// Core 3.10.2: deterministic typed walk, one bounded response window.
// Static facets carry no write capability. Every reused slot is cleared.
FUNCTION "FRK_ConfigRevision" : UDInt
{ S7_Optimized_Access := 'TRUE' }
VERSION : 0.1
VAR_INPUT
    Previous : UDInt;
END_VAR
VAR_TEMP
    Stamp : DTL;
    ResultCode : Int;
    Generation : ULInt;
END_VAR
BEGIN
    #FRK_ConfigRevision := #Previous + 1;
    #ResultCode := RD_SYS_T(OUT => #Stamp);
    IF #ResultCode = 0 THEN
        #Generation := LDT_TO_ULINT(DTL_TO_LDT(#Stamp)) / ULINT#1000000;
        #FRK_ConfigRevision := ULINT_TO_UDINT(#Generation MOD ULINT#4294967296);
    END_IF;
    IF #FRK_ConfigRevision = #Previous THEN #FRK_ConfigRevision := #Previous + 1; END_IF;
    IF #FRK_ConfigRevision = 0 THEN #FRK_ConfigRevision := 1; END_IF;
END_FUNCTION

FUNCTION "FRK_ConfigBegin" : Void
{ S7_Optimized_Access := 'TRUE' }
VERSION : 0.1
VAR_INPUT
    PageIndex : DInt;
    Revision : UDInt;
END_VAR
VAR_IN_OUT
    Cursor : "FRK_ConfigCursor";
    Page : "ST_ConfigPage";
END_VAR
VAR_TEMP
    Index : Int;
END_VAR
BEGIN
    #Cursor.Position := 0;
    #Cursor.First := 0;
    #Page.Revision := #Revision;
    #Page.PageIndex := 0;
    IF #PageIndex >= 0 AND #PageIndex <= 32767 THEN
        #Cursor.First := #PageIndex * 16;
        #Page.PageIndex := DINT_TO_INT(#PageIndex);
    END_IF;
    #Page.PageCount := 1;
    #Page.EntryCount := 0;
    "FRK_UnitScratch".EmptyConfigEntry.ValueType := 1;
    "FRK_UnitScratch".EmptyConfigEntry.Readable := TRUE;
    FOR #Index := 1 TO 16 DO
        #Page.Entries[#Index] := "FRK_UnitScratch".EmptyConfigEntry;
    END_FOR;
END_FUNCTION

FUNCTION "FRK_ConfigAppend" : Void
{ S7_Optimized_Access := 'TRUE' }
VERSION : 0.1
VAR_INPUT
    Scope : String;
    Item : String;
    ValueText : WString;
    ValueType : DInt;
    ReadLevel : DInt;
    Readable : Bool;
END_VAR
VAR_IN_OUT
    Cursor : "FRK_ConfigCursor";
    Page : "ST_ConfigPage";
END_VAR
VAR_TEMP
    Slot : DInt;
END_VAR
BEGIN
    #Slot := #Cursor.Position - #Cursor.First;
    #Cursor.Position := #Cursor.Position + 1;
    IF #Slot < 0 OR #Slot >= 16 THEN RETURN; END_IF;
    #Slot := #Slot + 1;
    #Page.Entries[#Slot].Scope := STRING_TO_WSTRING(#Scope);
    #Page.Entries[#Slot].Item := STRING_TO_WSTRING(#Item);
    #Page.Entries[#Slot].ValueType := #ValueType;
    #Page.Entries[#Slot].ReadLevel := #ReadLevel;
    #Page.Entries[#Slot].Readable := #Readable;
    IF #Readable THEN #Page.Entries[#Slot].ValueText := #ValueText; END_IF;
    #Page.EntryCount := DINT_TO_INT(#Slot);
END_FUNCTION

FUNCTION "FRK_ConfigFinish" : Void
{ S7_Optimized_Access := 'TRUE' }
VERSION : 0.1
VAR_IN_OUT
    Cursor : "FRK_ConfigCursor";
    Page : "ST_ConfigPage";
END_VAR
BEGIN
    #Page.PageCount := DINT_TO_INT((#Cursor.Position + 16 - 1) / 16);
    IF #Page.PageCount < 1 THEN #Page.PageCount := 1; END_IF;
END_FUNCTION

FUNCTION "FRK_ConfigCatalog" : Void
{ S7_Optimized_Access := 'TRUE' }
VERSION : 0.1
VAR_INPUT
    Scope : String;
    Count : Int;
    Catalog : Array[1..12] of "ST_CommandInfo";
    ReadLevel : DInt;
    Readable : Bool;
END_VAR
VAR_IN_OUT
    Cursor : "FRK_ConfigCursor";
    Page : "ST_ConfigPage";
END_VAR
VAR_TEMP
    Index : Int;
    IndexText : String[8];
    Prefix : String[254];
    Item : String[254];
END_VAR
BEGIN
    "FRK_ConfigAppend"(Scope := #Scope, Item := 'CatalogCount', ValueText := STRING_TO_WSTRING(INT_TO_STRING(#Count)), ValueType := 0, ReadLevel := #ReadLevel, Readable := #Readable, Cursor := #Cursor, Page := #Page);
    FOR #Index := 1 TO #Count DO
        IF #Index > 12 THEN EXIT; END_IF;
        #IndexText := INT_TO_STRING(#Index);
        IF #IndexText[1] = '+' THEN #IndexText := DELETE(IN := #IndexText, L := 1, P := 1); END_IF;
        #Prefix := CONCAT(IN1 := 'Catalog/Catalog[', IN2 := #IndexText);
        #Prefix := CONCAT(IN1 := #Prefix, IN2 := ']/');
        #Item := CONCAT(IN1 := #Prefix, IN2 := 'Value');
        "FRK_ConfigAppend"(Scope := #Scope, Item := #Item, ValueText := STRING_TO_WSTRING(DINT_TO_STRING(#Catalog[#Index].Value)), ValueType := 0, ReadLevel := #ReadLevel, Readable := #Readable, Cursor := #Cursor, Page := #Page);
        #Item := CONCAT(IN1 := #Prefix, IN2 := 'Label');
        "FRK_ConfigAppend"(Scope := #Scope, Item := #Item, ValueText := STRING_TO_WSTRING(#Catalog[#Index].Label), ValueType := 1, ReadLevel := #ReadLevel, Readable := #Readable, Cursor := #Cursor, Page := #Page);
        #Item := CONCAT(IN1 := #Prefix, IN2 := 'Style');
        "FRK_ConfigAppend"(Scope := #Scope, Item := #Item, ValueText := STRING_TO_WSTRING(DINT_TO_STRING(#Catalog[#Index].Style)), ValueType := 0, ReadLevel := #ReadLevel, Readable := #Readable, Cursor := #Cursor, Page := #Page);
    END_FOR;
END_FUNCTION

FUNCTION "FRK_ConfigUnit" : Void
{ S7_Optimized_Access := 'TRUE' }
VERSION : 0.1
VAR_INPUT
    Scope : String;
    Policy : Array[0..6] of "ST_ModePolicy";
    ModelCount : Int;
    ReadLevel : DInt;
    Readable : Bool;
END_VAR
VAR_IN_OUT
    Cursor : "FRK_ConfigCursor";
    Page : "ST_ConfigPage";
END_VAR
VAR_TEMP
    Index : Int;
    IndexText : String[8];
    Prefix : String[254];
    Item : String[254];
END_VAR
BEGIN
    "FRK_ConfigAppend"(Scope := #Scope, Item := 'CatalogCount', ValueText := WSTRING#'0', ValueType := 0, ReadLevel := #ReadLevel, Readable := #Readable, Cursor := #Cursor, Page := #Page);
    "FRK_ConfigAppend"(Scope := #Scope, Item := 'AvailableModelCount', ValueText := INT_TO_WSTRING(#ModelCount), ValueType := 0, ReadLevel := #ReadLevel, Readable := #Readable, Cursor := #Cursor, Page := #Page);
    FOR #Index := 0 TO 6 DO
        #IndexText := INT_TO_STRING(#Index);
        IF #IndexText[1] = '+' THEN #IndexText := DELETE(IN := #IndexText, L := 1, P := 1); END_IF;
        #Prefix := CONCAT(IN1 := 'ModePolicy/ModePolicy[', IN2 := #IndexText);
        #Prefix := CONCAT(IN1 := #Prefix, IN2 := ']/');
        #Item := CONCAT(IN1 := #Prefix, IN2 := 'Shield');
        "FRK_ConfigAppend"(Scope := #Scope, Item := #Item, ValueText := STRING_TO_WSTRING(DINT_TO_STRING(#Policy[#Index].Shield)), ValueType := 0, ReadLevel := #ReadLevel, Readable := #Readable, Cursor := #Cursor, Page := #Page);
        #Item := CONCAT(IN1 := #Prefix, IN2 := 'Style');
        "FRK_ConfigAppend"(Scope := #Scope, Item := #Item, ValueText := STRING_TO_WSTRING(DINT_TO_STRING(#Policy[#Index].Style)), ValueType := 0, ReadLevel := #ReadLevel, Readable := #Readable, Cursor := #Cursor, Page := #Page);
    END_FOR;
END_FUNCTION

// Core 8.3: one owning active list / closed ring, with optional event callback.
FUNCTION "FRK_AlarmNotify" : Void
{ S7_Optimized_Access := 'TRUE' }
VERSION : 0.1
VAR_INPUT
    Ev : "ST_AlarmEvent";
END_VAR
VAR_IN_OUT
    AlarmLog : "FRK_AlarmLog";
END_VAR
BEGIN
    RETURN; // No event sink supplied by the composition declaration.
END_FUNCTION

FUNCTION "FRK_AlarmRefresh" : Void
{ S7_Optimized_Access := 'TRUE' }
VERSION : 0.1
VAR_IN_OUT
    AlarmLog : "FRK_AlarmLog";
END_VAR
VAR_TEMP
    Index : Int;
END_VAR
BEGIN
    #AlarmLog.NActive := 0;
    #AlarmLog.Blocking := FALSE;
    FOR #Index := 1 TO 16 DO
        IF #AlarmLog.Active[#Index].State <> 0 THEN
            #AlarmLog.NActive := #AlarmLog.NActive + 1;
            IF #AlarmLog.Active[#Index].ResetClass = 1 THEN #AlarmLog.Blocking := TRUE; END_IF;
        END_IF;
    END_FOR;
    "FRK_AlarmRecoveryRefresh"(AlarmLog := #AlarmLog);
END_FUNCTION

FUNCTION "FRK_AlarmBegin" : Void
{ S7_Optimized_Access := 'TRUE' }
VERSION : 0.1
VAR_INPUT
    Startup : Bool;
END_VAR
VAR_IN_OUT
    AlarmLog : "FRK_AlarmLog";
END_VAR
VAR_TEMP
    Index : Int;
END_VAR
BEGIN
    FOR #Index := 1 TO 16 DO
        #AlarmLog.Touched[#Index] := FALSE;
        IF #Startup THEN
            #AlarmLog.Active[#Index] := "FRK_UnitScratch".EmptyEvent;
            #AlarmLog.Automatic[#Index] := FALSE;
            #AlarmLog.ComeMs[#Index] := 0;
        END_IF;
    END_FOR;
    IF #Startup THEN
        FOR #Index := 1 TO 64 DO #AlarmLog.Ring[#Index] := "FRK_UnitScratch".EmptyEvent; END_FOR;
        #AlarmLog.RingHead := 0;
        #AlarmLog.RingUsed := 0;
        #AlarmLog.Truncated := FALSE;
    END_IF;
    IF #Startup AND #AlarmLog.HistorySlot > 0 THEN "FRK_AlarmHistoryClear"(AlarmLog := #AlarmLog); END_IF;
    IF #Startup THEN "FRK_AlarmRecoveryClear"(AlarmLog := #AlarmLog); END_IF;
    "FRK_AlarmRefresh"(AlarmLog := #AlarmLog);
END_FUNCTION

FUNCTION "FRK_AlarmRaise" : Int
{ S7_Optimized_Access := 'TRUE' }
VERSION : 0.1
VAR_INPUT
    Diag : "ST_Diagnostic";
    ResetClass : DInt;
END_VAR
VAR_IN_OUT
    AlarmLog : "FRK_AlarmLog";
END_VAR
VAR_TEMP
    Slot : Int;
    Stamp : DTL;
    ResultCode : Int;
    Rational : "ST_Diagnostic";
END_VAR
BEGIN
    #FRK_AlarmRaise := 0;
    IF #ResetClass < 0 OR #ResetClass > 1
        OR #Diag.Severity < 0 OR #Diag.Severity > 2
        OR #Diag.Category < 0 OR #Diag.Category > 2
        OR #Diag.SourcePath = WSTRING#'' OR #Diag.Description = WSTRING#'' THEN RETURN; END_IF;
    #Slot := "FRK_AlarmRecoveryClaim"(AlarmLog := #AlarmLog, Diag := #Diag, ResetClass := #ResetClass); IF #Slot > 0 THEN #FRK_AlarmRaise := #Slot; RETURN; END_IF;
    FOR #Slot := 1 TO 16 DO
        IF #AlarmLog.Active[#Slot].State = 0 THEN
            #Rational := #Diag;
            "FRK_Rationalize"(Diag := #Rational);
            #AlarmLog.Active[#Slot] := "FRK_UnitScratch".EmptyEvent;
            #AlarmLog.Active[#Slot].ReasonCode := #Rational.ReasonCode;
            #AlarmLog.Active[#Slot].Description := #Rational.Description;
            #AlarmLog.Active[#Slot].SourcePath := #Rational.SourcePath;
            #AlarmLog.Active[#Slot].IoTag := #Rational.IoTag;
            #AlarmLog.Active[#Slot].IoAddress := #Rational.IoAddress;
            #AlarmLog.Active[#Slot].Severity := #Rational.Severity;
            #AlarmLog.Active[#Slot].Category := #Rational.Category;
            #AlarmLog.Active[#Slot].ResetClass := #ResetClass;
            #AlarmLog.Active[#Slot].State := 1;
            #AlarmLog.ComeMs[#Slot] := "FRK_Clock".NowMs;
            #AlarmLog.ElapsedBefore[#Slot] := 0; #AlarmLog.Recovering[#Slot] := FALSE;
            #AlarmLog.Automatic[#Slot] := FALSE;
            #AlarmLog.Touched[#Slot] := FALSE;
            #ResultCode := RD_SYS_T(OUT => #Stamp);
            IF #ResultCode = 0 THEN #AlarmLog.Active[#Slot].ComeAt := DTL_TO_LDT(#Stamp); END_IF;
            // The UTC source has no proven synchronization witness yet.
            #AlarmLog.Active[#Slot].ComeTimeSynchronized := FALSE;
            "FRK_AlarmRefresh"(AlarmLog := #AlarmLog);
            "FRK_AlarmRecoveryStore"(AlarmLog := #AlarmLog, EventSlot := #Slot);
            "FRK_DeliveryCapture"(AlarmLog := #AlarmLog, Ev := #AlarmLog.Active[#Slot]);
            "FRK_AlarmNotify"(AlarmLog := #AlarmLog, Ev := #AlarmLog.Active[#Slot]);
            #FRK_AlarmRaise := #Slot;
            RETURN;
        END_IF;
    END_FOR;
    IF NOT #AlarmLog.Truncated THEN
        #AlarmLog.Truncated := TRUE;
        "FRK_AlarmHistoryHeaderSave"(AlarmLog := #AlarmLog);
    END_IF;
END_FUNCTION

FUNCTION "FRK_AlarmClose" : Void
{ S7_Optimized_Access := 'TRUE' }
VERSION : 0.1
VAR_INPUT
    Slot : Int;
END_VAR
VAR_IN_OUT
    AlarmLog : "FRK_AlarmLog";
END_VAR
BEGIN
    IF #Slot < 1 OR #Slot > 16 THEN RETURN; END_IF;
    IF #AlarmLog.Active[#Slot].State = 0 THEN RETURN; END_IF;
    #AlarmLog.Active[#Slot].State := 0;
    "FRK_DeliveryCapture"(AlarmLog := #AlarmLog, Ev := #AlarmLog.Active[#Slot]);
    "FRK_AlarmRecoveryClosePrepare"(AlarmLog := #AlarmLog, EventSlot := #Slot);
    IF #AlarmLog.RingHead < 0 OR #AlarmLog.RingHead > 64 THEN #AlarmLog.RingHead := 0; END_IF;
    #AlarmLog.RingHead := (#AlarmLog.RingHead MOD 64) + 1;
    IF #AlarmLog.RingUsed >= 64 THEN #AlarmLog.Truncated := TRUE;
    ELSE #AlarmLog.RingUsed := #AlarmLog.RingUsed + 1; END_IF;
    #AlarmLog.Ring[#AlarmLog.RingHead] := #AlarmLog.Active[#Slot];
    "FRK_AlarmHistoryAppend"(AlarmLog := #AlarmLog);
    "FRK_AlarmRecoveryStore"(AlarmLog := #AlarmLog, EventSlot := #Slot);
    #AlarmLog.Automatic[#Slot] := FALSE;
    "FRK_AlarmRefresh"(AlarmLog := #AlarmLog);
    "FRK_AlarmNotify"(AlarmLog := #AlarmLog, Ev := #AlarmLog.Ring[#AlarmLog.RingHead]);
END_FUNCTION

FUNCTION "FRK_AlarmGone" : Bool
{ S7_Optimized_Access := 'TRUE' }
VERSION : 0.1
VAR_INPUT
    Slot : Int;
END_VAR
VAR_IN_OUT
    AlarmLog : "FRK_AlarmLog";
END_VAR
VAR_TEMP
    Span : UDInt;
    Stamp : DTL;
    ResultCode : Int;
END_VAR
BEGIN
    #FRK_AlarmGone := FALSE;
    IF #Slot < 1 OR #Slot > 16 THEN RETURN; END_IF;
    IF #AlarmLog.Active[#Slot].State <> 1 THEN RETURN; END_IF;
    #ResultCode := RD_SYS_T(OUT => #Stamp);
    IF #ResultCode = 0 THEN #AlarmLog.Active[#Slot].GoneAt := DTL_TO_LDT(#Stamp); END_IF;
    #AlarmLog.Active[#Slot].GoneTimeSynchronized := FALSE;
    #Span := "FRK_AlarmRecoveryElapsed"(AlarmLog := #AlarmLog, EventSlot := #Slot);
    #AlarmLog.Active[#Slot].Duration := DINT_TO_TIME(UDINT_TO_DINT(#Span));
    IF #AlarmLog.Active[#Slot].ResetClass = 0 THEN
        "FRK_AlarmClose"(AlarmLog := #AlarmLog, Slot := #Slot);
    ELSE
        #AlarmLog.Active[#Slot].State := 2;
        #AlarmLog.Automatic[#Slot] := FALSE;
        "FRK_AlarmRecoveryStore"(AlarmLog := #AlarmLog, EventSlot := #Slot);
    END_IF;
    #FRK_AlarmGone := TRUE;
END_FUNCTION

FUNCTION "FRK_AlarmOperatorReset" : Void
{ S7_Optimized_Access := 'TRUE' }
VERSION : 0.1
VAR_IN_OUT
    AlarmLog : "FRK_AlarmLog";
END_VAR
VAR_TEMP
    Slot : Int;
    Gone : Bool;
    Stamp : DTL;
    ResultCode : Int;
END_VAR
BEGIN
    FOR #Slot := 1 TO 16 DO
        IF #AlarmLog.Active[#Slot].State <> 0 AND #AlarmLog.Active[#Slot].ResetClass = 1 THEN
            IF #AlarmLog.Active[#Slot].State = 1 THEN #Gone := "FRK_AlarmGone"(AlarmLog := #AlarmLog, Slot := #Slot); END_IF;
            #ResultCode := RD_SYS_T(OUT => #Stamp);
            IF #ResultCode = 0 THEN #AlarmLog.Active[#Slot].ResetAt := DTL_TO_LDT(#Stamp); END_IF;
            #AlarmLog.Active[#Slot].ResetTimeSynchronized := FALSE;
            "FRK_AlarmClose"(AlarmLog := #AlarmLog, Slot := #Slot);
        END_IF;
    END_FOR;
END_FUNCTION

FUNCTION "FRK_AlarmMessage" : Void
{ S7_Optimized_Access := 'TRUE' }
VERSION : 0.1
VAR_INPUT
    Reason : DInt;
    Description : WString;
    SourcePath : WString;
END_VAR
VAR_IN_OUT
    AlarmLog : "FRK_AlarmLog";
END_VAR
VAR_TEMP
    Diag : "ST_Diagnostic";
    Slot : Int;
    Gone : Bool;
END_VAR
BEGIN
    #Diag := "FRK_UnitScratch".EmptyDiagnostic;
    #Diag.ReasonCode := #Reason;
    #Diag.Description := #Description;
    #Diag.SourcePath := #SourcePath;
    #Diag.Severity := 0;
    #Diag.Category := 2;
    #Slot := "FRK_AlarmRaise"(AlarmLog := #AlarmLog, Diag := #Diag, ResetClass := 0);
    IF #Slot > 0 THEN #Gone := "FRK_AlarmGone"(AlarmLog := #AlarmLog, Slot := #Slot); END_IF;
END_FUNCTION

FUNCTION "FRK_AlarmCapture" : Void
{ S7_Optimized_Access := 'TRUE' }
VERSION : 0.1
VAR_IN_OUT
    AlarmLog : "FRK_AlarmLog";
    Core : "FRK_Core";
    Status : "ST_ModuleStatus";
END_VAR
VAR_TEMP
    Slot : Int;
END_VAR
BEGIN
    #Slot := #Core.FaultSlot;
    IF #Slot < 1 OR #Slot > 16 THEN #Slot := 0;
    ELSIF NOT #AlarmLog.Automatic[#Slot] OR #AlarmLog.Active[#Slot].State <> 1
        OR #AlarmLog.Active[#Slot].SourcePath <> #Status.Diagnostic.SourcePath
        OR #AlarmLog.Active[#Slot].ReasonCode <> #Status.Diagnostic.ReasonCode
        OR #AlarmLog.Active[#Slot].Description <> #Status.Diagnostic.Description THEN #Slot := 0; END_IF;
    IF #Core.Exec = 3 AND NOT #Core.FaultHandled THEN
        IF #Slot = 0 THEN
            // Adopted first-outs share one active occurrence within this log.
            FOR #Slot := 1 TO 16 DO
                IF #AlarmLog.Automatic[#Slot] AND #AlarmLog.Active[#Slot].State = 1
                    AND #AlarmLog.Active[#Slot].SourcePath = #Status.Diagnostic.SourcePath
                    AND #AlarmLog.Active[#Slot].ReasonCode = #Status.Diagnostic.ReasonCode
                    AND #AlarmLog.Active[#Slot].Description = #Status.Diagnostic.Description THEN EXIT; END_IF;
            END_FOR;
            IF #Slot > 16 THEN #Slot := "FRK_AlarmRaise"(AlarmLog := #AlarmLog, Diag := #Status.Diagnostic, ResetClass := 1); END_IF;
        END_IF;
        IF #Slot > 0 THEN IF NOT #AlarmLog.Automatic[#Slot] THEN #AlarmLog.Automatic[#Slot] := TRUE; "FRK_AlarmRecoveryStore"(AlarmLog := #AlarmLog, EventSlot := #Slot); END_IF; #AlarmLog.Recovering[#Slot] := FALSE; #AlarmLog.Automatic[#Slot] := TRUE; #AlarmLog.Touched[#Slot] := TRUE; END_IF;
        #Core.FaultSlot := #Slot;
    ELSE
        #Core.FaultSlot := 0;
    END_IF;
END_FUNCTION

FUNCTION "FRK_AlarmEnd" : Void
{ S7_Optimized_Access := 'TRUE' }
VERSION : 0.1
VAR_IN_OUT
    AlarmLog : "FRK_AlarmLog";
END_VAR
VAR_TEMP
    Slot : Int;
    Gone : Bool;
END_VAR
BEGIN
    FOR #Slot := 1 TO 16 DO
        IF #AlarmLog.Automatic[#Slot] AND NOT #AlarmLog.Touched[#Slot] THEN #Gone := "FRK_AlarmGone"(AlarmLog := #AlarmLog, Slot := #Slot); END_IF;
    END_FOR;
END_FUNCTION

FUNCTION "FRK_AlarmTreeBlocking" : Bool
{ S7_Optimized_Access := 'TRUE' }
VERSION : 0.1
VAR_INPUT
    Owner : DInt;
END_VAR
VAR_TEMP
    Index : DInt;
    Ancestor : DInt;
    Depth : DInt;
END_VAR
BEGIN
    #FRK_AlarmTreeBlocking := TRUE;
    IF "FRK_Registry".Fault OR #Owner < 1 OR #Owner > "FRK_Registry".Count OR "FRK_Registry".Count > 4 THEN RETURN; END_IF;
    FOR #Index := 1 TO "FRK_Registry".Count DO
        IF "FRK_Registry".Rows[#Index].AlarmBlocking THEN
            #Ancestor := #Index;
            FOR #Depth := 1 TO 4 DO
                IF #Ancestor = #Owner THEN RETURN; END_IF;
                IF #Ancestor = 0 THEN EXIT; END_IF;
                IF #Ancestor < 1 OR #Ancestor > "FRK_Registry".Count THEN RETURN; END_IF;
                #Ancestor := "FRK_Registry".Rows[#Ancestor].Parent;
            END_FOR;
            IF #Depth > 4 AND #Ancestor <> 0 THEN RETURN; END_IF;
        END_IF;
    END_FOR;
    #FRK_AlarmTreeBlocking := FALSE;
END_FUNCTION

// Reference-1500 LOCAL_RETAIN: closed history only, keyed by actual Unit scope.
// No active alarms, commands, sessions or monotonic clocks are restored.
FUNCTION "FRK_AlarmHistoryIndex" : Int
{ S7_Optimized_Access := 'TRUE' }
VERSION : 0.1
VAR_INPUT
    Scope : String;
END_VAR
BEGIN
    #FRK_AlarmHistoryIndex := 0;
    IF #Scope = 'PressDemo' THEN #FRK_AlarmHistoryIndex := 1; RETURN; END_IF;
END_FUNCTION

FUNCTION "FRK_AlarmEventCrc" : DWord
{ S7_Optimized_Access := 'TRUE' }
VERSION : 0.1
VAR_INPUT
    Ev : "ST_AlarmEvent";
END_VAR
VAR_TEMP
    Work : DWord;
    Index : Int;
    Size : Int;
    Code : Word;
    Wide : LWord;
END_VAR
BEGIN
    #Work := DWORD#16#FFFFFFFF;
    #Work := "FRK_CrcNumber"(Previous := #Work, Value := DINT_TO_UDINT(#Ev.ReasonCode));
    #Size := LEN(#Ev.Description);
    #Work := "FRK_CrcNumber"(Previous := #Work, Value := INT_TO_UDINT(#Size));
    FOR #Index := 1 TO #Size DO
        #Code := WCHAR_TO_WORD(#Ev.Description[#Index]);
        #Work := "FRK_CrcByte"(Previous := #Work, Value := WORD_TO_BYTE(#Code));
        #Work := "FRK_CrcByte"(Previous := #Work, Value := WORD_TO_BYTE(SHR(IN := #Code, N := 8)));
    END_FOR;
    #Size := LEN(#Ev.SourcePath);
    #Work := "FRK_CrcNumber"(Previous := #Work, Value := INT_TO_UDINT(#Size));
    FOR #Index := 1 TO #Size DO
        #Code := WCHAR_TO_WORD(#Ev.SourcePath[#Index]);
        #Work := "FRK_CrcByte"(Previous := #Work, Value := WORD_TO_BYTE(#Code));
        #Work := "FRK_CrcByte"(Previous := #Work, Value := WORD_TO_BYTE(SHR(IN := #Code, N := 8)));
    END_FOR;
    #Size := LEN(#Ev.IoTag);
    #Work := "FRK_CrcNumber"(Previous := #Work, Value := INT_TO_UDINT(#Size));
    FOR #Index := 1 TO #Size DO
        #Work := "FRK_CrcByte"(Previous := #Work, Value := CHAR_TO_BYTE(#Ev.IoTag[#Index]));
    END_FOR;
    #Size := LEN(#Ev.IoAddress);
    #Work := "FRK_CrcNumber"(Previous := #Work, Value := INT_TO_UDINT(#Size));
    FOR #Index := 1 TO #Size DO
        #Work := "FRK_CrcByte"(Previous := #Work, Value := CHAR_TO_BYTE(#Ev.IoAddress[#Index]));
    END_FOR;
    #Work := "FRK_CrcNumber"(Previous := #Work, Value := DINT_TO_UDINT(#Ev.Severity));
    #Work := "FRK_CrcNumber"(Previous := #Work, Value := DINT_TO_UDINT(#Ev.Category));
    #Work := "FRK_CrcNumber"(Previous := #Work, Value := DINT_TO_UDINT(#Ev.ResetClass));
    #Work := "FRK_CrcNumber"(Previous := #Work, Value := DINT_TO_UDINT(#Ev.State));
    #Wide := LINT_TO_LWORD(LDT_TO_LINT(#Ev.ComeAt));
    #Work := "FRK_CrcNumber"(Previous := #Work, Value := DWORD_TO_UDINT(LWORD_TO_DWORD(#Wide)));
    #Work := "FRK_CrcNumber"(Previous := #Work, Value := DWORD_TO_UDINT(LWORD_TO_DWORD(SHR(IN := #Wide, N := 32))));
    #Wide := LINT_TO_LWORD(LDT_TO_LINT(#Ev.GoneAt));
    #Work := "FRK_CrcNumber"(Previous := #Work, Value := DWORD_TO_UDINT(LWORD_TO_DWORD(#Wide)));
    #Work := "FRK_CrcNumber"(Previous := #Work, Value := DWORD_TO_UDINT(LWORD_TO_DWORD(SHR(IN := #Wide, N := 32))));
    #Wide := LINT_TO_LWORD(LDT_TO_LINT(#Ev.ResetAt));
    #Work := "FRK_CrcNumber"(Previous := #Work, Value := DWORD_TO_UDINT(LWORD_TO_DWORD(#Wide)));
    #Work := "FRK_CrcNumber"(Previous := #Work, Value := DWORD_TO_UDINT(LWORD_TO_DWORD(SHR(IN := #Wide, N := 32))));
    #Work := "FRK_CrcNumber"(Previous := #Work, Value := DINT_TO_UDINT(TIME_TO_DINT(#Ev.Duration)));
    #Work := "FRK_CrcNumber"(Previous := #Work, Value := BOOL_TO_UDINT(#Ev.Shelved));
    #Wide := LINT_TO_LWORD(LDT_TO_LINT(#Ev.ShelvedUntil));
    #Work := "FRK_CrcNumber"(Previous := #Work, Value := DWORD_TO_UDINT(LWORD_TO_DWORD(#Wide)));
    #Work := "FRK_CrcNumber"(Previous := #Work, Value := DWORD_TO_UDINT(LWORD_TO_DWORD(SHR(IN := #Wide, N := 32))));
    #Work := "FRK_CrcNumber"(Previous := #Work, Value := BOOL_TO_UDINT(#Ev.ComeTimeSynchronized));
    #Work := "FRK_CrcNumber"(Previous := #Work, Value := BOOL_TO_UDINT(#Ev.GoneTimeSynchronized));
    #Work := "FRK_CrcNumber"(Previous := #Work, Value := BOOL_TO_UDINT(#Ev.ResetTimeSynchronized));
    #Work := "FRK_CrcNumber"(Previous := #Work, Value := BOOL_TO_UDINT(#Ev.ShelfTimeSynchronized));
    #FRK_AlarmEventCrc := NOT #Work;
END_FUNCTION

FUNCTION "FRK_AlarmHistoryHeaderCrc" : DWord
{ S7_Optimized_Access := 'TRUE' }
VERSION : 0.1
VAR_INPUT
    Slot : Int;
END_VAR
VAR_TEMP
    Work : DWord;
    Index : Int;
    Size : Int;
END_VAR
BEGIN
    #FRK_AlarmHistoryHeaderCrc := DWORD#0;
    IF #Slot < 1 OR #Slot > 1 THEN RETURN; END_IF;
    #Work := "FRK_CrcNumber"(Previous := DWORD#16#FFFFFFFF, Value := UINT_TO_UDINT("FRK_AlarmHistory".Rows[#Slot].SchemaVersion));
    #Size := LEN("FRK_AlarmHistory".Rows[#Slot].Scope);
    #Work := "FRK_CrcNumber"(Previous := #Work, Value := INT_TO_UDINT(#Size));
    FOR #Index := 1 TO #Size DO
        #Work := "FRK_CrcByte"(Previous := #Work, Value := CHAR_TO_BYTE("FRK_AlarmHistory".Rows[#Slot].Scope[#Index]));
    END_FOR;
    #Work := "FRK_CrcNumber"(Previous := #Work, Value := "FRK_AlarmHistory".Rows[#Slot].Generation);
    #Work := "FRK_CrcNumber"(Previous := #Work, Value := INT_TO_UDINT("FRK_AlarmHistory".Rows[#Slot].RingHead));
    #Work := "FRK_CrcNumber"(Previous := #Work, Value := INT_TO_UDINT("FRK_AlarmHistory".Rows[#Slot].RingUsed));
    #Work := "FRK_CrcNumber"(Previous := #Work, Value := BOOL_TO_UDINT("FRK_AlarmHistory".Rows[#Slot].Truncated));
    FOR #Index := 1 TO 64 DO
        #Work := "FRK_CrcNumber"(Previous := #Work, Value := DWORD_TO_UDINT("FRK_AlarmHistory".Rows[#Slot].EventCrc[#Index]));
    END_FOR;
    #FRK_AlarmHistoryHeaderCrc := NOT #Work;
END_FUNCTION

FUNCTION "FRK_AlarmHistoryHeaderSave" : Void
{ S7_Optimized_Access := 'TRUE' }
VERSION : 0.1
VAR_IN_OUT
    AlarmLog : "FRK_AlarmLog";
END_VAR
VAR_TEMP
    Slot : Int;
END_VAR
BEGIN
    #Slot := #AlarmLog.HistorySlot;
    IF #Slot < 1 OR #Slot > 1 THEN RETURN; END_IF;
    "FRK_AlarmHistory".Rows[#Slot].SchemaVersion := 1;
    "FRK_AlarmHistory".Rows[#Slot].Generation := "FRK_AccessNext"(Previous := "FRK_AlarmHistory".Rows[#Slot].Generation);
    "FRK_AlarmHistory".Rows[#Slot].RingHead := #AlarmLog.RingHead;
    "FRK_AlarmHistory".Rows[#Slot].RingUsed := #AlarmLog.RingUsed;
    "FRK_AlarmHistory".Rows[#Slot].Truncated := #AlarmLog.Truncated;
    "FRK_AlarmHistory".Rows[#Slot].Checksum := "FRK_AlarmHistoryHeaderCrc"(Slot := #Slot);
    "FRK_AlarmHistory".Commissioned[#Slot] := TRUE;
END_FUNCTION

FUNCTION "FRK_AlarmHistoryClear" : Void
{ S7_Optimized_Access := 'TRUE' }
VERSION : 0.1
VAR_IN_OUT
    AlarmLog : "FRK_AlarmLog";
END_VAR
VAR_TEMP
    Index : Int;
    Slot : Int;
END_VAR
BEGIN
    #Slot := #AlarmLog.HistorySlot;
    IF #Slot < 1 OR #Slot > 1 THEN RETURN; END_IF;
    FOR #Index := 1 TO 64 DO
        "FRK_AlarmHistory".Rows[#Slot].Ring[#Index] := "FRK_UnitScratch".EmptyEvent;
        "FRK_AlarmHistory".Rows[#Slot].EventCrc[#Index] := DWORD#0;
    END_FOR;
    "FRK_AlarmHistoryHeaderSave"(AlarmLog := #AlarmLog);
END_FUNCTION

FUNCTION "FRK_AlarmHistoryAppend" : Void
{ S7_Optimized_Access := 'TRUE' }
VERSION : 0.1
VAR_IN_OUT
    AlarmLog : "FRK_AlarmLog";
END_VAR
VAR_TEMP
    Slot : Int;
    Head : Int;
END_VAR
BEGIN
    #Slot := #AlarmLog.HistorySlot;
    #Head := #AlarmLog.RingHead;
    IF #Slot < 1 OR #Slot > 1 OR #Head < 1 OR #Head > 64 THEN RETURN; END_IF;
    "FRK_AlarmHistory".Rows[#Slot].Ring[#Head] := #AlarmLog.Ring[#Head];
    "FRK_AlarmHistory".Rows[#Slot].EventCrc[#Head] := "FRK_AlarmEventCrc"(Ev := #AlarmLog.Ring[#Head]);
    "FRK_AlarmHistoryHeaderSave"(AlarmLog := #AlarmLog);
END_FUNCTION

FUNCTION "FRK_AlarmHistoryBoot" : Void
{ S7_Optimized_Access := 'TRUE' }
VERSION : 0.1
VAR_INPUT
    Startup : Bool;
    Scope : String;
END_VAR
VAR_IN_OUT
    AlarmLog : "FRK_AlarmLog";
END_VAR
VAR_TEMP
    Slot : Int;
    Index : Int;
    Used : Int;
    Head : Int;
    Valid : Bool;
END_VAR
BEGIN
    IF NOT #Startup THEN RETURN; END_IF;
    #Slot := "FRK_AlarmHistoryIndex"(Scope := #Scope);
    #AlarmLog.HistorySlot := #Slot;
    IF #Slot < 1 OR #Slot > 1 THEN RETURN; END_IF;
    IF NOT "FRK_AlarmHistory".Commissioned[#Slot]
        AND "FRK_AlarmHistory".Rows[#Slot].SchemaVersion = 0
        AND "FRK_AlarmHistory".Rows[#Slot].Generation = 0
        AND "FRK_AlarmHistory".Rows[#Slot].Scope = ''
        AND "FRK_AlarmHistory".Rows[#Slot].Checksum = DWORD#0 THEN
        "FRK_AlarmHistory".Rows[#Slot].Scope := #Scope;
        "FRK_AlarmHistoryClear"(AlarmLog := #AlarmLog);
        RETURN;
    END_IF;
    #Used := "FRK_AlarmHistory".Rows[#Slot].RingUsed;
    #Head := "FRK_AlarmHistory".Rows[#Slot].RingHead;
    #Valid := "FRK_AlarmHistory".Rows[#Slot].SchemaVersion = 1
        AND "FRK_AlarmHistory".Rows[#Slot].Scope = #Scope
        AND "FRK_AlarmHistory".Rows[#Slot].Generation <> 0
        AND #Used >= 0 AND #Used <= 64
        AND #Head >= 0 AND #Head <= 64
        AND ((#Used = 0 AND #Head = 0) OR (#Used > 0 AND #Head > 0))
        AND (#Used = 64 OR #Head = #Used);
    IF #Valid THEN #Valid := "FRK_AlarmHistory".Rows[#Slot].Checksum = "FRK_AlarmHistoryHeaderCrc"(Slot := #Slot); END_IF;
    IF #Valid THEN
        FOR #Index := 1 TO #Used DO
            IF "FRK_AlarmHistory".Rows[#Slot].Ring[#Index].State <> 0
                OR "FRK_AlarmHistory".Rows[#Slot].Ring[#Index].ResetClass < 0
                OR "FRK_AlarmHistory".Rows[#Slot].Ring[#Index].ResetClass > 1
                OR "FRK_AlarmHistory".Rows[#Slot].Ring[#Index].Severity < 0
                OR "FRK_AlarmHistory".Rows[#Slot].Ring[#Index].Severity > 2
                OR "FRK_AlarmHistory".Rows[#Slot].Ring[#Index].Category < 0
                OR "FRK_AlarmHistory".Rows[#Slot].Ring[#Index].Category > 2
                OR "FRK_AlarmHistory".Rows[#Slot].Ring[#Index].SourcePath = WSTRING#''
                OR "FRK_AlarmHistory".Rows[#Slot].Ring[#Index].Description = WSTRING#''
                OR "FRK_AlarmHistory".Rows[#Slot].Ring[#Index].Duration < T#0ms
                OR "FRK_AlarmHistory".Rows[#Slot].EventCrc[#Index] <> "FRK_AlarmEventCrc"(Ev := "FRK_AlarmHistory".Rows[#Slot].Ring[#Index]) THEN
                #Valid := FALSE;
                EXIT;
            END_IF;
        END_FOR;
    END_IF;
    IF #Valid THEN
        FOR #Index := 1 TO #Used DO #AlarmLog.Ring[#Index] := "FRK_AlarmHistory".Rows[#Slot].Ring[#Index]; END_FOR;
        #AlarmLog.RingHead := #Head;
        #AlarmLog.RingUsed := #Used;
        #AlarmLog.Truncated := "FRK_AlarmHistory".Rows[#Slot].Truncated;
    ELSE
        // Reject the whole image. The same public loss marker covers overflow
        // and rejected history; do not present a partial, apparently complete log.
        #AlarmLog.Truncated := TRUE;
        "FRK_AlarmHistory".Rows[#Slot].Scope := #Scope;
        "FRK_AlarmHistoryClear"(AlarmLog := #AlarmLog);
    END_IF;
END_FUNCTION

// Binding-local opt-in recovery of manual-reset latches. Commands remain volatile.
FUNCTION "FRK_AlarmRecoveryIndex" : Int
{ S7_Optimized_Access := 'TRUE' }
VERSION : 0.1
VAR_INPUT
    Scope : String;
END_VAR
BEGIN
    #FRK_AlarmRecoveryIndex := 0;
    IF #Scope = 'PressDemo' THEN #FRK_AlarmRecoveryIndex := 1; RETURN; END_IF;
END_FUNCTION

FUNCTION "FRK_AlarmRecoveryScope" : String
{ S7_Optimized_Access := 'TRUE' }
VERSION : 0.1
VAR_INPUT
    Slot : Int;
END_VAR
BEGIN
    CASE #Slot OF
        1: #FRK_AlarmRecoveryScope := 'PressDemo';
        ELSE #FRK_AlarmRecoveryScope := '';
    END_CASE;
END_FUNCTION

FUNCTION "FRK_AlarmRecoveryPrepare" : Void
{ S7_Optimized_Access := 'TRUE' }
VERSION : 0.1
VAR_INPUT
    Startup : Bool;
END_VAR
VAR_TEMP
    Slot : Int;
END_VAR
BEGIN
    IF NOT #Startup THEN RETURN; END_IF;
    // All selected descendants are conservative until their owning frame restores.
    FOR #Slot := 1 TO 1 DO
        "FRK_AlarmRecoveryRuntime".Ready[#Slot] := FALSE;
        "FRK_AlarmRecoveryRuntime".Blocked[#Slot] := TRUE;
    END_FOR;
END_FUNCTION

FUNCTION "FRK_AlarmRecoveryTreeBlocking" : Bool
{ S7_Optimized_Access := 'TRUE' }
VERSION : 0.1
VAR_INPUT
    Scope : String;
END_VAR
VAR_TEMP
    Slot : Int;
    Expected : String[80];
    Prefix : String[80];
END_VAR
BEGIN
    #FRK_AlarmRecoveryTreeBlocking := FALSE;
    #Prefix := CONCAT(IN1 := #Scope, IN2 := '.');
    FOR #Slot := 1 TO 1 DO
        #Expected := "FRK_AlarmRecoveryScope"(Slot := #Slot);
        IF #Expected = #Scope OR LEFT(IN := #Expected, L := LEN(#Prefix)) = #Prefix THEN
            IF NOT "FRK_AlarmRecoveryRuntime".Ready[#Slot] OR "FRK_AlarmRecoveryRuntime".Blocked[#Slot] THEN
                #FRK_AlarmRecoveryTreeBlocking := TRUE; RETURN;
            END_IF;
        END_IF;
    END_FOR;
END_FUNCTION

FUNCTION "FRK_AlarmRecoveryRefresh" : Void
{ S7_Optimized_Access := 'TRUE' }
VERSION : 0.1
VAR_IN_OUT
    AlarmLog : "FRK_AlarmLog";
END_VAR
BEGIN
    IF #AlarmLog.RecoverySlot < 1 OR #AlarmLog.RecoverySlot > 1 THEN RETURN; END_IF;
    "FRK_AlarmRecoveryRuntime".Blocked[#AlarmLog.RecoverySlot] := #AlarmLog.Blocking;
END_FUNCTION

FUNCTION "FRK_AlarmRecoveryElapsed" : UDInt
{ S7_Optimized_Access := 'TRUE' }
VERSION : 0.1
VAR_INPUT
    EventSlot : Int;
END_VAR
VAR_IN_OUT
    AlarmLog : "FRK_AlarmLog";
END_VAR
VAR_TEMP
    Span : UDInt;
END_VAR
BEGIN
    #FRK_AlarmRecoveryElapsed := 0;
    IF #EventSlot < 1 OR #EventSlot > 16 THEN RETURN; END_IF;
    #Span := "FRK_Elapsed"(NewMs := "FRK_Clock".NowMs, OldMs := #AlarmLog.ComeMs[#EventSlot]);
    IF #Span > 2147483647 - #AlarmLog.ElapsedBefore[#EventSlot] THEN #Span := 2147483647;
    ELSE #Span := #Span + #AlarmLog.ElapsedBefore[#EventSlot]; END_IF;
    #FRK_AlarmRecoveryElapsed := #Span;
END_FUNCTION

FUNCTION "FRK_AlarmRecoveryTimeCrc" : DWord
{ S7_Optimized_Access := 'TRUE' }
VERSION : 0.1
VAR_INPUT
    Slot : Int;
    EventSlot : Int;
    Value : UDInt;
    EventCrc : DWord;
END_VAR
VAR_TEMP
    Work : DWord;
END_VAR
BEGIN
    #Work := "FRK_CrcNumber"(Previous := DWORD#16#FFFFFFFF, Value := INT_TO_UDINT(#Slot));
    #Work := "FRK_CrcNumber"(Previous := #Work, Value := INT_TO_UDINT(#EventSlot));
    #Work := "FRK_CrcNumber"(Previous := #Work, Value := DWORD_TO_UDINT(#EventCrc));
    #Work := "FRK_CrcNumber"(Previous := #Work, Value := #Value);
    #FRK_AlarmRecoveryTimeCrc := NOT #Work;
END_FUNCTION

FUNCTION "FRK_AlarmRecoveryHeaderCrc" : DWord
{ S7_Optimized_Access := 'TRUE' }
VERSION : 0.1
VAR_INPUT
    Slot : Int;
END_VAR
VAR_TEMP
    Work : DWord;
    Index : Int;
    Size : Int;
END_VAR
BEGIN
    #FRK_AlarmRecoveryHeaderCrc := DWORD#0;
    IF #Slot < 1 OR #Slot > 1 THEN RETURN; END_IF;
    #Work := "FRK_CrcNumber"(Previous := DWORD#16#FFFFFFFF, Value := UINT_TO_UDINT("FRK_AlarmRecovery".Rows[#Slot].SchemaVersion));
    #Size := LEN("FRK_AlarmRecovery".Rows[#Slot].Scope);
    #Work := "FRK_CrcNumber"(Previous := #Work, Value := INT_TO_UDINT(#Size));
    FOR #Index := 1 TO #Size DO
        #Work := "FRK_CrcByte"(Previous := #Work, Value := CHAR_TO_BYTE("FRK_AlarmRecovery".Rows[#Slot].Scope[#Index]));
    END_FOR;
    #Work := "FRK_CrcNumber"(Previous := #Work, Value := "FRK_AlarmRecovery".Rows[#Slot].Generation);
    FOR #Index := 1 TO 16 DO
        #Work := "FRK_CrcNumber"(Previous := #Work, Value := DWORD_TO_UDINT("FRK_AlarmRecovery".Rows[#Slot].EventCrc[#Index]));
        #Work := "FRK_CrcNumber"(Previous := #Work, Value := BOOL_TO_UDINT("FRK_AlarmRecovery".Rows[#Slot].Automatic[#Index]));
    END_FOR;
    #Work := "FRK_CrcNumber"(Previous := #Work, Value := INT_TO_UDINT("FRK_AlarmRecovery".Rows[#Slot].PendingSlot));
    #Work := "FRK_CrcNumber"(Previous := #Work, Value := DWORD_TO_UDINT("FRK_AlarmRecovery".Rows[#Slot].PendingCrc));
    #Work := "FRK_CrcNumber"(Previous := #Work, Value := INT_TO_UDINT("FRK_AlarmRecovery".Rows[#Slot].PendingHead));
    #Work := "FRK_CrcNumber"(Previous := #Work, Value := "FRK_AlarmRecovery".Rows[#Slot].PendingHistoryGeneration);
    #FRK_AlarmRecoveryHeaderCrc := NOT #Work;
END_FUNCTION

FUNCTION "FRK_AlarmRecoveryHeaderSave" : Void
{ S7_Optimized_Access := 'TRUE' }
VERSION : 0.1
VAR_INPUT
    Slot : Int;
END_VAR
BEGIN
    IF #Slot < 1 OR #Slot > 1 THEN RETURN; END_IF;
    "FRK_AlarmRecovery".Rows[#Slot].SchemaVersion := 2;
    "FRK_AlarmRecovery".Rows[#Slot].Generation := "FRK_AccessNext"(Previous := "FRK_AlarmRecovery".Rows[#Slot].Generation);
    "FRK_AlarmRecovery".Rows[#Slot].Checksum := "FRK_AlarmRecoveryHeaderCrc"(Slot := #Slot);
    "FRK_AlarmRecovery".Commissioned[#Slot] := TRUE;
END_FUNCTION

FUNCTION "FRK_AlarmRecoveryClear" : Void
{ S7_Optimized_Access := 'TRUE' }
VERSION : 0.1
VAR_IN_OUT
    AlarmLog : "FRK_AlarmLog";
END_VAR
VAR_TEMP
    Slot : Int;
    Index : Int;
END_VAR
BEGIN
    #Slot := #AlarmLog.RecoverySlot;
    IF #Slot < 1 OR #Slot > 1 THEN RETURN; END_IF;
    FOR #Index := 1 TO 16 DO
        "FRK_AlarmRecovery".Rows[#Slot].Active[#Index] := "FRK_UnitScratch".EmptyEvent;
        "FRK_AlarmRecovery".Rows[#Slot].EventCrc[#Index] := DWORD#0;
        "FRK_AlarmRecovery".Rows[#Slot].Automatic[#Index] := FALSE;
        "FRK_AlarmRecovery".Rows[#Slot].Elapsed[#Index] := 0;
        "FRK_AlarmRecovery".Rows[#Slot].TimeCrc[#Index] := DWORD#0;
        "FRK_AlarmRecovery".Rows[#Slot].ElapsedAlt[#Index] := 0;
        "FRK_AlarmRecovery".Rows[#Slot].TimeCrcAlt[#Index] := DWORD#0;
        "FRK_AlarmRecovery".Rows[#Slot].TimeBank[#Index] := FALSE;
        #AlarmLog.ElapsedBefore[#Index] := 0;
        #AlarmLog.Recovering[#Index] := FALSE;
    END_FOR;
    "FRK_AlarmRecovery".Rows[#Slot].PendingSlot := 0;
    "FRK_AlarmRecovery".Rows[#Slot].PendingClosed := "FRK_UnitScratch".EmptyEvent;
    "FRK_AlarmRecovery".Rows[#Slot].PendingCrc := DWORD#0;
    "FRK_AlarmRecovery".Rows[#Slot].PendingHead := 0;
    "FRK_AlarmRecovery".Rows[#Slot].PendingHistoryGeneration := 0;
    "FRK_AlarmRecoveryHeaderSave"(Slot := #Slot);
END_FUNCTION

FUNCTION "FRK_AlarmRecoveryStore" : Void
{ S7_Optimized_Access := 'TRUE' }
VERSION : 0.1
VAR_INPUT
    EventSlot : Int;
END_VAR
VAR_IN_OUT
    AlarmLog : "FRK_AlarmLog";
END_VAR
VAR_TEMP
    Slot : Int;
    Span : UDInt;
END_VAR
BEGIN
    #Slot := #AlarmLog.RecoverySlot;
    IF #Slot < 1 OR #Slot > 1 OR #EventSlot < 1 OR #EventSlot > 16 THEN RETURN; END_IF;
    IF #AlarmLog.Active[#EventSlot].State <> 0 AND #AlarmLog.Active[#EventSlot].ResetClass = 1 THEN
        "FRK_AlarmRecovery".Rows[#Slot].Active[#EventSlot] := #AlarmLog.Active[#EventSlot];
        "FRK_AlarmRecovery".Rows[#Slot].EventCrc[#EventSlot] := "FRK_AlarmEventCrc"(Ev := #AlarmLog.Active[#EventSlot]);
        "FRK_AlarmRecovery".Rows[#Slot].Automatic[#EventSlot] := #AlarmLog.Automatic[#EventSlot];
        IF #AlarmLog.Active[#EventSlot].State = 1 THEN #Span := "FRK_AlarmRecoveryElapsed"(AlarmLog := #AlarmLog, EventSlot := #EventSlot);
        ELSE #Span := DINT_TO_UDINT(TIME_TO_DINT(#AlarmLog.Active[#EventSlot].Duration)); END_IF;
        "FRK_AlarmRecovery".Rows[#Slot].Elapsed[#EventSlot] := #Span;
        "FRK_AlarmRecovery".Rows[#Slot].TimeCrc[#EventSlot] := "FRK_AlarmRecoveryTimeCrc"(Slot := #Slot, EventSlot := #EventSlot, Value := #Span, EventCrc := "FRK_AlarmRecovery".Rows[#Slot].EventCrc[#EventSlot]);
        "FRK_AlarmRecovery".Rows[#Slot].ElapsedAlt[#EventSlot] := #Span;
        "FRK_AlarmRecovery".Rows[#Slot].TimeCrcAlt[#EventSlot] := "FRK_AlarmRecovery".Rows[#Slot].TimeCrc[#EventSlot];
        "FRK_AlarmRecovery".Rows[#Slot].TimeBank[#EventSlot] := FALSE;
    ELSE
        IF "FRK_AlarmRecovery".Rows[#Slot].Active[#EventSlot].State = 0 AND "FRK_AlarmRecovery".Rows[#Slot].PendingSlot <> #EventSlot THEN RETURN; END_IF;
        "FRK_AlarmRecovery".Rows[#Slot].Active[#EventSlot] := "FRK_UnitScratch".EmptyEvent;
        "FRK_AlarmRecovery".Rows[#Slot].EventCrc[#EventSlot] := DWORD#0;
        "FRK_AlarmRecovery".Rows[#Slot].Automatic[#EventSlot] := FALSE;
        "FRK_AlarmRecovery".Rows[#Slot].Elapsed[#EventSlot] := 0;
        "FRK_AlarmRecovery".Rows[#Slot].TimeCrc[#EventSlot] := DWORD#0;
        "FRK_AlarmRecovery".Rows[#Slot].ElapsedAlt[#EventSlot] := 0;
        "FRK_AlarmRecovery".Rows[#Slot].TimeCrcAlt[#EventSlot] := DWORD#0;
        "FRK_AlarmRecovery".Rows[#Slot].TimeBank[#EventSlot] := FALSE;
        #AlarmLog.ElapsedBefore[#EventSlot] := 0;
        #AlarmLog.Recovering[#EventSlot] := FALSE;
    END_IF;
    IF "FRK_AlarmRecovery".Rows[#Slot].PendingSlot = #EventSlot THEN
        "FRK_AlarmRecovery".Rows[#Slot].PendingSlot := 0;
        "FRK_AlarmRecovery".Rows[#Slot].PendingClosed := "FRK_UnitScratch".EmptyEvent;
        "FRK_AlarmRecovery".Rows[#Slot].PendingCrc := DWORD#0;
        "FRK_AlarmRecovery".Rows[#Slot].PendingHead := 0;
        "FRK_AlarmRecovery".Rows[#Slot].PendingHistoryGeneration := 0;
    END_IF;
    "FRK_AlarmRecoveryHeaderSave"(Slot := #Slot);
END_FUNCTION

FUNCTION "FRK_AlarmRecoveryCheckpointRead" : Void
{ S7_Optimized_Access := 'TRUE' }
VERSION : 0.1
VAR_INPUT
    Slot : Int;
    EventSlot : Int;
END_VAR
VAR_OUTPUT
    Elapsed : UDInt;
    Checksum : DWord;
END_VAR
BEGIN
    #Elapsed := 0; #Checksum := DWORD#0;
    IF #Slot < 1 OR #Slot > 1 OR #EventSlot < 1 OR #EventSlot > 16 THEN RETURN; END_IF;
    IF "FRK_AlarmRecovery".Rows[#Slot].TimeBank[#EventSlot] THEN
        #Elapsed := "FRK_AlarmRecovery".Rows[#Slot].ElapsedAlt[#EventSlot];
        #Checksum := "FRK_AlarmRecovery".Rows[#Slot].TimeCrcAlt[#EventSlot];
    ELSE
        #Elapsed := "FRK_AlarmRecovery".Rows[#Slot].Elapsed[#EventSlot];
        #Checksum := "FRK_AlarmRecovery".Rows[#Slot].TimeCrc[#EventSlot];
    END_IF;
END_FUNCTION

FUNCTION "FRK_AlarmRecoveryTick" : Void
{ S7_Optimized_Access := 'TRUE' }
VERSION : 0.1
VAR_IN_OUT
    AlarmLog : "FRK_AlarmLog";
END_VAR
VAR_TEMP
    Slot : Int;
    Index : Int;
    Span : UDInt;
    Saved : UDInt;
    SavedCrc : DWord;
    Work : DWord;
END_VAR
BEGIN
    #Slot := #AlarmLog.RecoverySlot;
    IF #Slot < 1 OR #Slot > 1 THEN RETURN; END_IF;
    FOR #Index := 1 TO 16 DO
        IF #AlarmLog.Active[#Index].State = 1 AND #AlarmLog.Active[#Index].ResetClass = 1 THEN
            #Span := "FRK_AlarmRecoveryElapsed"(AlarmLog := #AlarmLog, EventSlot := #Index);
            "FRK_AlarmRecoveryCheckpointRead"(Slot := #Slot, EventSlot := #Index, Elapsed => #Saved, Checksum => #SavedCrc);
            IF #Saved <> #Span THEN
                #Work := "FRK_AlarmRecoveryTimeCrc"(Slot := #Slot, EventSlot := #Index, Value := #Span, EventCrc := "FRK_AlarmRecovery".Rows[#Slot].EventCrc[#Index]);
                IF "FRK_AlarmRecovery".Rows[#Slot].TimeBank[#Index] THEN
                    "FRK_AlarmRecovery".Rows[#Slot].Elapsed[#Index] := #Span;
                    "FRK_AlarmRecovery".Rows[#Slot].TimeCrc[#Index] := #Work;
                ELSE
                    "FRK_AlarmRecovery".Rows[#Slot].ElapsedAlt[#Index] := #Span;
                    "FRK_AlarmRecovery".Rows[#Slot].TimeCrcAlt[#Index] := #Work;
                END_IF;
                "FRK_AlarmRecovery".Rows[#Slot].TimeBank[#Index] := NOT "FRK_AlarmRecovery".Rows[#Slot].TimeBank[#Index];
            END_IF;
        END_IF;
    END_FOR;
END_FUNCTION

FUNCTION "FRK_AlarmRecoveryClaim" : Int
{ S7_Optimized_Access := 'TRUE' }
VERSION : 0.1
VAR_INPUT
    Diag : "ST_Diagnostic";
    ResetClass : DInt;
END_VAR
VAR_IN_OUT
    AlarmLog : "FRK_AlarmLog";
END_VAR
VAR_TEMP
    Slot : Int;
END_VAR
BEGIN
    #FRK_AlarmRecoveryClaim := 0;
    IF #ResetClass <> 1 THEN RETURN; END_IF;
    FOR #Slot := 1 TO 16 DO
        IF #AlarmLog.Recovering[#Slot] AND #AlarmLog.Active[#Slot].State = 1
            AND #AlarmLog.Active[#Slot].ReasonCode = #Diag.ReasonCode
            AND #AlarmLog.Active[#Slot].Description = #Diag.Description
            AND #AlarmLog.Active[#Slot].SourcePath = #Diag.SourcePath THEN
            #AlarmLog.Recovering[#Slot] := FALSE;
            #FRK_AlarmRecoveryClaim := #Slot; RETURN;
        END_IF;
    END_FOR;
END_FUNCTION

FUNCTION "FRK_AlarmRecoveryClosePrepare" : Void
{ S7_Optimized_Access := 'TRUE' }
VERSION : 0.1
VAR_INPUT
    EventSlot : Int;
END_VAR
VAR_IN_OUT
    AlarmLog : "FRK_AlarmLog";
END_VAR
VAR_TEMP
    Slot : Int;
END_VAR
BEGIN
    #Slot := #AlarmLog.RecoverySlot;
    IF #Slot < 1 OR #Slot > 1 OR #EventSlot < 1 OR #EventSlot > 16 THEN RETURN; END_IF;
    IF #AlarmLog.Active[#EventSlot].ResetClass <> 1 THEN RETURN; END_IF;
    "FRK_AlarmRecovery".Rows[#Slot].PendingSlot := #EventSlot;
    "FRK_AlarmRecovery".Rows[#Slot].PendingClosed := #AlarmLog.Active[#EventSlot];
    "FRK_AlarmRecovery".Rows[#Slot].PendingCrc := "FRK_AlarmEventCrc"(Ev := #AlarmLog.Active[#EventSlot]);
    "FRK_AlarmRecovery".Rows[#Slot].PendingHead := (#AlarmLog.RingHead MOD 64) + 1;
    "FRK_AlarmRecovery".Rows[#Slot].PendingHistoryGeneration := "FRK_AccessNext"(Previous := "FRK_AlarmHistory".Rows[#AlarmLog.HistorySlot].Generation);
    "FRK_AlarmRecoveryHeaderSave"(Slot := #Slot);
END_FUNCTION

FUNCTION "FRK_AlarmRecoveryEventValid" : Bool
{ S7_Optimized_Access := 'TRUE' }
VERSION : 0.1
VAR_INPUT
    Ev : "ST_AlarmEvent";
END_VAR
BEGIN
    #FRK_AlarmRecoveryEventValid := #Ev.ResetClass = 1
        AND #Ev.Severity >= 0 AND #Ev.Severity <= 2
        AND #Ev.Category >= 0 AND #Ev.Category <= 2
        AND #Ev.SourcePath <> WSTRING#'' AND #Ev.Description <> WSTRING#'' AND #Ev.ReasonCode > 0 AND #Ev.Duration >= T#0ms;
END_FUNCTION

FUNCTION "FRK_AlarmRecoveryBoot" : Void
{ S7_Optimized_Access := 'TRUE' }
VERSION : 0.1
VAR_INPUT
    Startup : Bool;
    Scope : String;
END_VAR
VAR_IN_OUT
    AlarmLog : "FRK_AlarmLog";
END_VAR
VAR_TEMP
    Slot : Int;
    Index : Int;
    Pending : Int;
    Head : Int;
    Valid : Bool;
    ClosedPresent : Bool;
    LossSlot : Int;
    Diag : "ST_Diagnostic";
    SavedElapsed : UDInt;
    SavedCrc : DWord;
END_VAR
BEGIN
    IF NOT #Startup THEN RETURN; END_IF;
    #Slot := "FRK_AlarmRecoveryIndex"(Scope := #Scope);
    #AlarmLog.RecoverySlot := #Slot;
    IF #Slot < 1 OR #Slot > 1 THEN RETURN; END_IF;
    IF NOT "FRK_AlarmRecovery".Commissioned[#Slot] AND "FRK_AlarmRecovery".Rows[#Slot].SchemaVersion = 0
        AND "FRK_AlarmRecovery".Rows[#Slot].Generation = 0 AND "FRK_AlarmRecovery".Rows[#Slot].Scope = '' AND "FRK_AlarmRecovery".Rows[#Slot].Checksum = DWORD#0 THEN
        "FRK_AlarmRecovery".Rows[#Slot].Scope := #Scope;
        "FRK_AlarmRecoveryClear"(AlarmLog := #AlarmLog);
        "FRK_AlarmRecoveryRuntime".Ready[#Slot] := TRUE;
        "FRK_AlarmRefresh"(AlarmLog := #AlarmLog);
        RETURN;
    END_IF;
    #Valid := "FRK_AlarmRecovery".Rows[#Slot].SchemaVersion = 2 AND "FRK_AlarmRecovery".Rows[#Slot].Scope = #Scope
        AND "FRK_AlarmRecovery".Rows[#Slot].Generation <> 0;
    IF #Valid THEN #Valid := "FRK_AlarmRecovery".Rows[#Slot].Checksum = "FRK_AlarmRecoveryHeaderCrc"(Slot := #Slot); END_IF;
    IF #Valid THEN
        FOR #Index := 1 TO 16 DO
            "FRK_AlarmRecoveryCheckpointRead"(Slot := #Slot, EventSlot := #Index, Elapsed => #SavedElapsed, Checksum => #SavedCrc);
            IF "FRK_AlarmRecovery".Rows[#Slot].Active[#Index].State = 0 THEN
                IF "FRK_AlarmRecovery".Rows[#Slot].EventCrc[#Index] <> DWORD#0 OR #SavedElapsed <> 0
                    OR #SavedCrc <> DWORD#0 OR "FRK_AlarmRecovery".Rows[#Slot].Automatic[#Index] THEN #Valid := FALSE; EXIT; END_IF;
            ELSE
                IF NOT "FRK_AlarmRecoveryEventValid"(Ev := "FRK_AlarmRecovery".Rows[#Slot].Active[#Index])
                    OR ("FRK_AlarmRecovery".Rows[#Slot].Active[#Index].State <> 1 AND "FRK_AlarmRecovery".Rows[#Slot].Active[#Index].State <> 2)
                    OR "FRK_AlarmRecovery".Rows[#Slot].EventCrc[#Index] <> "FRK_AlarmEventCrc"(Ev := "FRK_AlarmRecovery".Rows[#Slot].Active[#Index])
                    OR #SavedElapsed > 2147483647
                    OR #SavedCrc <> "FRK_AlarmRecoveryTimeCrc"(Slot := #Slot, EventSlot := #Index, Value := #SavedElapsed, EventCrc := "FRK_AlarmRecovery".Rows[#Slot].EventCrc[#Index]) THEN #Valid := FALSE; EXIT; END_IF;
                IF "FRK_AlarmRecovery".Rows[#Slot].Active[#Index].State = 2
                    AND ("FRK_AlarmRecovery".Rows[#Slot].Automatic[#Index] OR #SavedElapsed <> DINT_TO_UDINT(TIME_TO_DINT("FRK_AlarmRecovery".Rows[#Slot].Active[#Index].Duration))) THEN #Valid := FALSE; EXIT; END_IF;
            END_IF;
        END_FOR;
    END_IF;
    #Pending := "FRK_AlarmRecovery".Rows[#Slot].PendingSlot;
    IF #Valid THEN
        IF #Pending < 0 OR #Pending > 16 THEN #Valid := FALSE;
        ELSIF #Pending = 0 THEN
            IF "FRK_AlarmRecovery".Rows[#Slot].PendingCrc <> DWORD#0 OR "FRK_AlarmRecovery".Rows[#Slot].PendingHead <> 0 OR "FRK_AlarmRecovery".Rows[#Slot].PendingHistoryGeneration <> 0 THEN #Valid := FALSE; END_IF;
        ELSE
            #Valid := "FRK_AlarmRecoveryEventValid"(Ev := "FRK_AlarmRecovery".Rows[#Slot].PendingClosed)
                AND "FRK_AlarmRecovery".Rows[#Slot].PendingClosed.State = 0
                AND "FRK_AlarmRecovery".Rows[#Slot].PendingCrc = "FRK_AlarmEventCrc"(Ev := "FRK_AlarmRecovery".Rows[#Slot].PendingClosed)
                AND "FRK_AlarmRecovery".Rows[#Slot].PendingHead >= 1 AND "FRK_AlarmRecovery".Rows[#Slot].PendingHead <= 64
                AND "FRK_AlarmRecovery".Rows[#Slot].PendingHistoryGeneration <> 0
                AND "FRK_AlarmRecovery".Rows[#Slot].Active[#Pending].State <> 0
                AND "FRK_AlarmRecovery".Rows[#Slot].PendingClosed.ReasonCode = "FRK_AlarmRecovery".Rows[#Slot].Active[#Pending].ReasonCode
                AND "FRK_AlarmRecovery".Rows[#Slot].PendingClosed.SourcePath = "FRK_AlarmRecovery".Rows[#Slot].Active[#Pending].SourcePath
                AND "FRK_AlarmRecovery".Rows[#Slot].PendingClosed.Description = "FRK_AlarmRecovery".Rows[#Slot].Active[#Pending].Description
                AND "FRK_AlarmRecovery".Rows[#Slot].PendingClosed.ComeAt = "FRK_AlarmRecovery".Rows[#Slot].Active[#Pending].ComeAt;
        END_IF;
    END_IF;
    IF NOT #Valid THEN
        // Unknown prior manual-reset latches fail closed until one deliberate reset.
        #AlarmLog.Truncated := TRUE;
        "FRK_AlarmHistoryHeaderSave"(AlarmLog := #AlarmLog);
        "FRK_AlarmRecovery".Rows[#Slot].Scope := #Scope;
        "FRK_AlarmRecoveryClear"(AlarmLog := #AlarmLog);
        #Diag := "FRK_UnitScratch".EmptyDiagnostic;
        #Diag.ReasonCode := 11001;
        #Diag.Description := WSTRING#'std.error.alarmRestoreLost';
        #Diag.SourcePath := STRING_TO_WSTRING(#Scope);
        #Diag.Severity := 2; #Diag.Category := 2;
        #LossSlot := "FRK_AlarmRaise"(AlarmLog := #AlarmLog, Diag := #Diag, ResetClass := 1);
    ELSE
        FOR #Index := 1 TO 16 DO
            "FRK_AlarmRecoveryCheckpointRead"(Slot := #Slot, EventSlot := #Index, Elapsed => #SavedElapsed, Checksum => #SavedCrc);
            IF "FRK_AlarmRecovery".Rows[#Slot].Active[#Index].State <> 0 THEN
                #AlarmLog.Active[#Index] := "FRK_AlarmRecovery".Rows[#Slot].Active[#Index];
                #AlarmLog.Automatic[#Index] := "FRK_AlarmRecovery".Rows[#Slot].Automatic[#Index];
                #AlarmLog.Recovering[#Index] := #AlarmLog.Active[#Index].State = 1;
                #AlarmLog.ComeMs[#Index] := "FRK_Clock".NowMs;
                IF #AlarmLog.Active[#Index].State = 1 THEN #AlarmLog.ElapsedBefore[#Index] := #SavedElapsed; END_IF;
            END_IF;
        END_FOR;
        IF #Pending > 0 THEN
            #Head := "FRK_AlarmRecovery".Rows[#Slot].PendingHead;
            #ClosedPresent := "FRK_AlarmHistory".Rows[#AlarmLog.HistorySlot].Generation = "FRK_AlarmRecovery".Rows[#Slot].PendingHistoryGeneration
                AND #AlarmLog.RingHead = #Head
                AND "FRK_AlarmHistory".Rows[#AlarmLog.HistorySlot].EventCrc[#Head] = "FRK_AlarmRecovery".Rows[#Slot].PendingCrc;
            IF NOT #ClosedPresent THEN
                #AlarmLog.RingHead := (#AlarmLog.RingHead MOD 64) + 1;
                IF #AlarmLog.RingUsed < 64 THEN #AlarmLog.RingUsed := #AlarmLog.RingUsed + 1; ELSE #AlarmLog.Truncated := TRUE; END_IF;
                #AlarmLog.Ring[#AlarmLog.RingHead] := "FRK_AlarmRecovery".Rows[#Slot].PendingClosed;
                "FRK_AlarmHistoryAppend"(AlarmLog := #AlarmLog);
            END_IF;
            #AlarmLog.Active[#Pending] := "FRK_UnitScratch".EmptyEvent;
            #AlarmLog.Automatic[#Pending] := FALSE;
            "FRK_AlarmRecoveryStore"(AlarmLog := #AlarmLog, EventSlot := #Pending);
        END_IF;
    END_IF;
    "FRK_AlarmRecoveryRuntime".Ready[#Slot] := TRUE;
    "FRK_AlarmRefresh"(AlarmLog := #AlarmLog);
END_FUNCTION

// Optional Core 8.3 sink adapter. FIFO ownership is private; delivery receipts
// use the existing root commit mailbox and never modify alarm/control state.
FUNCTION "FRK_DeliveryIndex" : Int
{ S7_Optimized_Access := 'TRUE' }
VERSION : 0.1
VAR_INPUT
    Scope : String;
END_VAR
BEGIN
    #FRK_DeliveryIndex := 0;
    IF #Scope = 'PressDemo' THEN #FRK_DeliveryIndex := 1; RETURN; END_IF;
END_FUNCTION

FUNCTION "FRK_DeliveryRootIndex" : Int
{ S7_Optimized_Access := 'TRUE' }
VERSION : 0.1
VAR_INPUT
    RootScope : String;
END_VAR
BEGIN
    #FRK_DeliveryRootIndex := 0;
    IF #RootScope = 'PressDemo' THEN #FRK_DeliveryRootIndex := 1; RETURN; END_IF;
END_FUNCTION

FUNCTION "FRK_DeliveryMailbox" : Void
{ S7_Optimized_Access := 'TRUE' }
VERSION : 0.1
VAR_INPUT
    RootScope : String;
    Access : "FRK_Access";
END_VAR
VAR_IN_OUT
    AlarmLog : "FRK_AlarmLog";
END_VAR
VAR_TEMP
    Slot : Int;
    SequenceBefore : UDInt;
    Receipt : "FRK_DeliveryReceipt";
    Request : "ST_HmiRequest";
    Accepted : Bool;
    What : WString[160];
END_VAR
BEGIN
    #Slot := "FRK_DeliveryRootIndex"(RootScope := #RootScope);
    IF #Slot < 1 OR #Slot > 1 THEN RETURN; END_IF;
    "FRK_EventDeliveryReceipt".Roots[#Slot] := #RootScope;
    #SequenceBefore := "FRK_EventDeliveryReceipt".Request[#Slot].Sequence;
    IF #SequenceBefore = 0 OR #SequenceBefore = "FRK_EventDeliveryRuntime".SeenReceipt[#Slot] THEN RETURN; END_IF;
    #Receipt := "FRK_EventDeliveryReceipt".Request[#Slot];
    IF #SequenceBefore <> "FRK_EventDeliveryReceipt".Request[#Slot].Sequence THEN RETURN; END_IF;
    #Request.TargetPath := STRING_TO_WSTRING(#Receipt.TargetPath);
    #Request.NameValue := #Receipt.Token;
    #Request.DurationMs := #Receipt.Checksum;
    #Request.Kind := 10001;
    #Request.BoolValue := #Receipt.DiscardLost;
    IF #Receipt.DiscardLost THEN
        #Request.Kind := 10002;
        #Request.NameValue := "FRK_DeliveryNumber"(Value := #Receipt.Epoch);
        #Request.TextValue := STRING_TO_WSTRING(#Receipt.StreamId);
    END_IF;
    #Accepted := FALSE;
    IF #Receipt.SchemaVersion = 1 THEN #Accepted := "FRK_DeliveryRequest"(RootScope := #RootScope, Request := #Request, Access := #Access); END_IF;
    "FRK_EventDeliveryRuntime".SeenReceipt[#Slot] := #SequenceBefore;
    // Audit metadata receipts locally, without creating work to acknowledge the
    // acknowledgement. The operator session's idle time is not refreshed.
    #What := WSTRING#'std.audit.accessDenied';
    IF #Accepted THEN #What := WSTRING#'std.audit.operatorAction'; END_IF;
    #What := CONCAT(IN1 := #What, IN2 := WSTRING#' eventDelivery=');
    #What := CONCAT(IN1 := #What, IN2 := DINT_TO_WSTRING(#Request.Kind));
    #AlarmLog.DeliveryMuted := TRUE;
    "FRK_AccessAudit"(AlarmLog := #AlarmLog, What := #What, Who := #Access.CurrentUser, SourcePath := STRING_TO_WSTRING(#RootScope));
    #AlarmLog.DeliveryMuted := FALSE;
    "FRK_EventDeliveryReceipt".Response[#Slot].SchemaVersion := 1;
    "FRK_EventDeliveryReceipt".Response[#Slot].Accepted := #Accepted;
    "FRK_EventDeliveryReceipt".Response[#Slot].AckSequence := #SequenceBefore;
END_FUNCTION

FUNCTION "FRK_DeliveryStatus" : Void
{ S7_Optimized_Access := 'TRUE' }
VERSION : 0.1
VAR_INPUT
    Scope : String;
END_VAR
VAR_IN_OUT
    AlarmLog : "FRK_AlarmLog";
END_VAR
VAR_TEMP
    Slot : Int;
    EventSlot : Int;
    Gone : Bool;
    Diag : "ST_Diagnostic";
END_VAR
BEGIN
    #Slot := #AlarmLog.DeliverySlot;
    IF #Slot < 1 OR #Slot > 1 THEN RETURN; END_IF;
    #EventSlot := #AlarmLog.DeliveryLossSlot;
    IF #EventSlot < 1 OR #EventSlot > 16 THEN #EventSlot := 0;
    ELSIF #AlarmLog.Active[#EventSlot].State <> 1
        OR #AlarmLog.Active[#EventSlot].ReasonCode <> 11002
        OR #AlarmLog.Active[#EventSlot].SourcePath <> STRING_TO_WSTRING(#Scope) THEN #EventSlot := 0; END_IF;
    IF NOT "FRK_EventDeliveryRuntime".Valid[#Slot] THEN
        IF #EventSlot = 0 THEN
            #Diag := "FRK_UnitScratch".EmptyDiagnostic;
            #Diag.ReasonCode := 11002;
            #Diag.Description := WSTRING#'std.error.eventDeliveryRestoreLost';
            #Diag.SourcePath := STRING_TO_WSTRING(#Scope);
            #Diag.Severity := 0;
            #Diag.Category := 2;
            #EventSlot := "FRK_AlarmRaise"(AlarmLog := #AlarmLog, Diag := #Diag, ResetClass := 0);
        END_IF;
        #AlarmLog.DeliveryLossSlot := #EventSlot;
    ELSE
        IF #EventSlot > 0 THEN #Gone := "FRK_AlarmGone"(AlarmLog := #AlarmLog, Slot := #EventSlot); END_IF;
        #AlarmLog.DeliveryLossSlot := 0;
    END_IF;
END_FUNCTION

FUNCTION "FRK_DeliveryScope" : String
{ S7_Optimized_Access := 'TRUE' }
VERSION : 0.1
VAR_INPUT
    Slot : Int;
END_VAR
BEGIN
    #FRK_DeliveryScope := '';
    CASE #Slot OF
        1: #FRK_DeliveryScope := 'PressDemo';
        ELSE RETURN;
    END_CASE;
END_FUNCTION

FUNCTION "FRK_DeliveryAnchorCrc" : DWord
{ S7_Optimized_Access := 'TRUE' }
VERSION : 0.1
VAR_INPUT
    Slot : Int;
END_VAR
VAR_TEMP
    Work : DWord;
    Index : Int;
END_VAR
BEGIN
    #FRK_DeliveryAnchorCrc := DWORD#0;
    IF #Slot < 1 OR #Slot > 1 THEN RETURN; END_IF;
    #Work := "FRK_CrcNumber"(Previous := DWORD#16#FFFFFFFF, Value := UINT_TO_UDINT("FRK_EventDeliveryStore".Anchors[#Slot].SchemaVersion));
    FOR #Index := 1 TO LEN("FRK_EventDeliveryStore".Anchors[#Slot].Scope) DO
        #Work := "FRK_CrcByte"(Previous := #Work, Value := CHAR_TO_BYTE("FRK_EventDeliveryStore".Anchors[#Slot].Scope[#Index]));
    END_FOR;
    #Work := "FRK_CrcByte"(Previous := #Work, Value := BYTE#0);
    FOR #Index := 1 TO LEN("FRK_EventDeliveryStore".Anchors[#Slot].StreamId) DO
        #Work := "FRK_CrcByte"(Previous := #Work, Value := CHAR_TO_BYTE("FRK_EventDeliveryStore".Anchors[#Slot].StreamId[#Index]));
    END_FOR;
    #Work := "FRK_CrcNumber"(Previous := #Work, Value := "FRK_EventDeliveryStore".Anchors[#Slot].Epoch);
    #FRK_DeliveryAnchorCrc := NOT #Work;
END_FUNCTION

FUNCTION "FRK_DeliveryHeaderCrc" : DWord
{ S7_Optimized_Access := 'TRUE' }
VERSION : 0.1
VAR_INPUT
    Slot : Int;
END_VAR
VAR_TEMP
    Work : DWord;
END_VAR
BEGIN
    #FRK_DeliveryHeaderCrc := DWORD#0;
    IF #Slot < 1 OR #Slot > 1 THEN RETURN; END_IF;
    #Work := "FRK_CrcNumber"(Previous := DWORD#16#FFFFFFFF, Value := UINT_TO_UDINT("FRK_EventDeliveryStore".Images[#Slot].SchemaVersion));
    #Work := "FRK_CrcNumber"(Previous := #Work, Value := "FRK_EventDeliveryStore".Images[#Slot].Epoch);
    #Work := "FRK_CrcNumber"(Previous := #Work, Value := "FRK_EventDeliveryStore".Images[#Slot].Revision);
    #Work := "FRK_CrcNumber"(Previous := #Work, Value := "FRK_EventDeliveryStore".Images[#Slot].NextSequence);
    #Work := "FRK_CrcNumber"(Previous := #Work, Value := INT_TO_UDINT("FRK_EventDeliveryStore".Images[#Slot].Head));
    #Work := "FRK_CrcNumber"(Previous := #Work, Value := INT_TO_UDINT("FRK_EventDeliveryStore".Images[#Slot].Count));
    #Work := "FRK_CrcNumber"(Previous := #Work, Value := BOOL_TO_UDINT("FRK_EventDeliveryStore".Images[#Slot].Overflow));
    #Work := "FRK_CrcNumber"(Previous := #Work, Value := "FRK_EventDeliveryStore".Images[#Slot].Dropped);
    #FRK_DeliveryHeaderCrc := NOT #Work;
END_FUNCTION

FUNCTION "FRK_DeliveryRowCrc" : DWord
{ S7_Optimized_Access := 'TRUE' }
VERSION : 0.1
VAR_INPUT
    Sequence : UDInt;
    Ev : "ST_AlarmEvent";
END_VAR
BEGIN
    #FRK_DeliveryRowCrc := "FRK_CrcNumber"(Previous := "FRK_AlarmEventCrc"(Ev := #Ev), Value := #Sequence);
END_FUNCTION

FUNCTION "FRK_DeliveryNumber" : String
{ S7_Optimized_Access := 'TRUE' }
VERSION : 0.1
VAR_INPUT
    Value : UDInt;
END_VAR
VAR_TEMP
    Text : String[12];
END_VAR
BEGIN
    #Text := UDINT_TO_STRING(#Value);
    IF LEFT(IN := #Text, L := 1) = '+' THEN #Text := RIGHT(IN := #Text, L := LEN(#Text) - 1); END_IF;
    #FRK_DeliveryNumber := #Text;
END_FUNCTION

FUNCTION "FRK_DeliveryToken" : String
{ S7_Optimized_Access := 'TRUE' }
VERSION : 0.1
VAR_INPUT
    Slot : Int;
    Sequence : UDInt;
END_VAR
VAR_TEMP
    Work : String[160];
END_VAR
BEGIN
    #FRK_DeliveryToken := '';
    IF #Slot < 1 OR #Slot > 1 THEN RETURN; END_IF;
    #Work := CONCAT(IN1 := "FRK_EventDeliveryStore".Anchors[#Slot].StreamId, IN2 := '/');
    #Work := CONCAT(IN1 := #Work, IN2 := "FRK_EventDeliveryStore".Anchors[#Slot].Scope);
    #Work := CONCAT(IN1 := #Work, IN2 := '/');
    #Work := CONCAT(IN1 := #Work, IN2 := "FRK_DeliveryNumber"(Value := "FRK_EventDeliveryStore".Anchors[#Slot].Epoch));
    #Work := CONCAT(IN1 := #Work, IN2 := '/');
    #FRK_DeliveryToken := CONCAT(IN1 := #Work, IN2 := "FRK_DeliveryNumber"(Value := #Sequence));
END_FUNCTION

FUNCTION "FRK_DeliveryPublish" : Void
{ S7_Optimized_Access := 'TRUE' }
VERSION : 0.1
VAR_INPUT
    Slot : Int;
END_VAR
VAR_TEMP
    Head : Int;
END_VAR
BEGIN
    IF #Slot < 1 OR #Slot > 1 THEN RETURN; END_IF;
    // Copy event text only on a lifecycle change; never every scan.
    IF "FRK_EventDeliveryRuntime".PublishedRevision[#Slot] = "FRK_EventDeliveryStore".Images[#Slot].Revision
        AND "FRK_EventDeliveryView".Rows[#Slot].SchemaVersion = 1 THEN RETURN; END_IF;
    "FRK_EventDeliveryView".Rows[#Slot].SchemaVersion := 1;
    "FRK_EventDeliveryView".Rows[#Slot].Scope := "FRK_DeliveryScope"(Slot := #Slot);
    "FRK_EventDeliveryView".Rows[#Slot].StreamId := '6c62c9b6-57d9-41b5-b689-e0540f642b31';
    "FRK_EventDeliveryView".Rows[#Slot].Capacity := 32;
    "FRK_EventDeliveryView".Rows[#Slot].AnchorValid := "FRK_EventDeliveryRuntime".AnchorValid[#Slot];
    "FRK_EventDeliveryView".Rows[#Slot].RestoreLost := NOT "FRK_EventDeliveryRuntime".Valid[#Slot];
    "FRK_EventDeliveryView".Rows[#Slot].Pending := 0;
    "FRK_EventDeliveryView".Rows[#Slot].Token := '';
    "FRK_EventDeliveryView".Rows[#Slot].Checksum := 0;
    "FRK_EventDeliveryView".Rows[#Slot].Ev := "FRK_UnitScratch".EmptyEvent;
    IF "FRK_EventDeliveryRuntime".AnchorValid[#Slot] THEN "FRK_EventDeliveryView".Rows[#Slot].Epoch := "FRK_EventDeliveryStore".Anchors[#Slot].Epoch; END_IF;
    IF "FRK_EventDeliveryRuntime".Valid[#Slot] THEN
        "FRK_EventDeliveryView".Rows[#Slot].Pending := "FRK_EventDeliveryStore".Images[#Slot].Count;
        "FRK_EventDeliveryView".Rows[#Slot].Overflow := "FRK_EventDeliveryStore".Images[#Slot].Overflow;
        "FRK_EventDeliveryView".Rows[#Slot].Dropped := "FRK_EventDeliveryStore".Images[#Slot].Dropped;
        #Head := "FRK_EventDeliveryStore".Images[#Slot].Head;
        IF "FRK_EventDeliveryStore".Images[#Slot].Count > 0 AND #Head >= 1 AND #Head <= 32 THEN
            "FRK_EventDeliveryView".Rows[#Slot].Token := "FRK_DeliveryToken"(Slot := #Slot, Sequence := "FRK_EventDeliveryStore".Images[#Slot].Entries[#Head].Sequence);
            "FRK_EventDeliveryView".Rows[#Slot].Checksum := DWORD_TO_UDINT("FRK_EventDeliveryStore".Images[#Slot].Entries[#Head].Checksum);
            "FRK_EventDeliveryView".Rows[#Slot].Ev := "FRK_EventDeliveryStore".Images[#Slot].Entries[#Head].Ev;
        END_IF;
    ELSE
        "FRK_EventDeliveryView".Rows[#Slot].Overflow := TRUE;
        "FRK_EventDeliveryView".Rows[#Slot].Dropped := 0;
    END_IF;
    "FRK_EventDeliveryRuntime".PublishedRevision[#Slot] := "FRK_EventDeliveryStore".Images[#Slot].Revision;
END_FUNCTION

FUNCTION "FRK_DeliverySave" : Void
{ S7_Optimized_Access := 'TRUE' }
VERSION : 0.1
VAR_INPUT
    Slot : Int;
END_VAR
BEGIN
    IF #Slot < 1 OR #Slot > 1 THEN RETURN; END_IF;
    "FRK_EventDeliveryStore".Images[#Slot].Revision := "FRK_ConfigRevision"(Previous := "FRK_EventDeliveryStore".Images[#Slot].Revision);
    "FRK_EventDeliveryStore".Images[#Slot].Checksum := "FRK_DeliveryHeaderCrc"(Slot := #Slot);
    "FRK_EventDeliveryRuntime".PublishedRevision[#Slot] := 0;
    "FRK_DeliveryPublish"(Slot := #Slot);
END_FUNCTION

FUNCTION "FRK_DeliveryInitialize" : Void
{ S7_Optimized_Access := 'TRUE' }
VERSION : 0.1
VAR_INPUT
    Slot : Int;
    Discarded : Bool;
END_VAR
VAR_TEMP
    Index : Int;
END_VAR
BEGIN
    IF #Slot < 1 OR #Slot > 1 THEN RETURN; END_IF;
    "FRK_EventDeliveryStore".Images[#Slot].SchemaVersion := 1;
    "FRK_EventDeliveryStore".Images[#Slot].Epoch := "FRK_EventDeliveryStore".Anchors[#Slot].Epoch;
    "FRK_EventDeliveryStore".Images[#Slot].Revision := 0;
    "FRK_EventDeliveryStore".Images[#Slot].NextSequence := 0;
    "FRK_EventDeliveryStore".Images[#Slot].Head := 1;
    "FRK_EventDeliveryStore".Images[#Slot].Count := 0;
    "FRK_EventDeliveryStore".Images[#Slot].Overflow := #Discarded;
    "FRK_EventDeliveryStore".Images[#Slot].Dropped := 0;
    FOR #Index := 1 TO 32 DO
        "FRK_EventDeliveryStore".Images[#Slot].Entries[#Index].Sequence := 0;
        "FRK_EventDeliveryStore".Images[#Slot].Entries[#Index].Checksum := DWORD#0;
        "FRK_EventDeliveryStore".Images[#Slot].Entries[#Index].Ev := "FRK_UnitScratch".EmptyEvent;
    END_FOR;
    "FRK_EventDeliveryRuntime".Valid[#Slot] := TRUE;
    "FRK_DeliverySave"(Slot := #Slot);
    "FRK_EventDeliveryStore".Commissioned[#Slot] := TRUE;
END_FUNCTION

FUNCTION "FRK_DeliveryBoot" : Void
{ S7_Optimized_Access := 'TRUE' }
VERSION : 0.1
VAR_INPUT
    Scope : String;
    Startup : Bool;
END_VAR
VAR_IN_OUT
    AlarmLog : "FRK_AlarmLog";
END_VAR
VAR_TEMP
    Slot : Int;
    Index : Int;
    Position : Int;
    Previous : UDInt;
    Valid : Bool;
    AnchorOk : Bool;
    Ev : "ST_AlarmEvent";
END_VAR
BEGIN
    IF NOT #Startup THEN RETURN; END_IF;
    #Slot := "FRK_DeliveryIndex"(Scope := #Scope);
    #AlarmLog.DeliverySlot := #Slot;
    IF #Slot < 1 OR #Slot > 1 THEN RETURN; END_IF;
    "FRK_EventDeliveryRuntime".PublishedRevision[#Slot] := 0;
    "FRK_EventDeliveryView".Rows[#Slot].SchemaVersion := 0;
    IF NOT "FRK_EventDeliveryStore".Commissioned[#Slot]
        AND "FRK_EventDeliveryStore".Anchors[#Slot].SchemaVersion = 0
        AND "FRK_EventDeliveryStore".Anchors[#Slot].Epoch = 0
        AND "FRK_EventDeliveryStore".Anchors[#Slot].Scope = ''
        AND "FRK_EventDeliveryStore".Anchors[#Slot].StreamId = ''
        AND "FRK_EventDeliveryStore".Anchors[#Slot].Checksum = DWORD#0
        AND "FRK_EventDeliveryStore".Images[#Slot].SchemaVersion = 0
        AND "FRK_EventDeliveryStore".Images[#Slot].Revision = 0
        AND "FRK_EventDeliveryStore".Images[#Slot].Checksum = DWORD#0 THEN
        "FRK_EventDeliveryStore".Anchors[#Slot].SchemaVersion := 1;
        "FRK_EventDeliveryStore".Anchors[#Slot].Scope := #Scope;
        "FRK_EventDeliveryStore".Anchors[#Slot].StreamId := '6c62c9b6-57d9-41b5-b689-e0540f642b31';
        "FRK_EventDeliveryStore".Anchors[#Slot].Epoch := 1;
        "FRK_EventDeliveryStore".Anchors[#Slot].Checksum := "FRK_DeliveryAnchorCrc"(Slot := #Slot);
        "FRK_EventDeliveryRuntime".AnchorValid[#Slot] := TRUE;
        "FRK_DeliveryInitialize"(Slot := #Slot, Discarded := FALSE);
        RETURN;
    END_IF;
    #AnchorOk := "FRK_EventDeliveryStore".Commissioned[#Slot]
        AND "FRK_EventDeliveryStore".Anchors[#Slot].SchemaVersion = 1
        AND "FRK_EventDeliveryStore".Anchors[#Slot].Scope = #Scope
        AND "FRK_EventDeliveryStore".Anchors[#Slot].StreamId = '6c62c9b6-57d9-41b5-b689-e0540f642b31'
        AND "FRK_EventDeliveryStore".Anchors[#Slot].Epoch > 0;
    IF #AnchorOk THEN #AnchorOk := "FRK_EventDeliveryStore".Anchors[#Slot].Checksum = "FRK_DeliveryAnchorCrc"(Slot := #Slot); END_IF;
    "FRK_EventDeliveryRuntime".AnchorValid[#Slot] := #AnchorOk;
    #Valid := #AnchorOk AND "FRK_EventDeliveryStore".Images[#Slot].SchemaVersion = 1
        AND "FRK_EventDeliveryStore".Images[#Slot].Epoch = "FRK_EventDeliveryStore".Anchors[#Slot].Epoch
        AND "FRK_EventDeliveryStore".Images[#Slot].Revision > 0
        AND "FRK_EventDeliveryStore".Images[#Slot].Head >= 1 AND "FRK_EventDeliveryStore".Images[#Slot].Head <= 32
        AND "FRK_EventDeliveryStore".Images[#Slot].Count >= 0 AND "FRK_EventDeliveryStore".Images[#Slot].Count <= 32;
    IF #Valid THEN #Valid := "FRK_EventDeliveryStore".Images[#Slot].Checksum = "FRK_DeliveryHeaderCrc"(Slot := #Slot); END_IF;
    #Previous := 0;
    IF #Valid THEN
        FOR #Index := 0 TO "FRK_EventDeliveryStore".Images[#Slot].Count - 1 DO
            #Position := (("FRK_EventDeliveryStore".Images[#Slot].Head - 1 + #Index) MOD 32) + 1;
            #Ev := "FRK_EventDeliveryStore".Images[#Slot].Entries[#Position].Ev;
            #Valid := "FRK_EventDeliveryStore".Images[#Slot].Entries[#Position].Sequence > #Previous
                AND "FRK_EventDeliveryStore".Images[#Slot].Entries[#Position].Sequence <= "FRK_EventDeliveryStore".Images[#Slot].NextSequence
                AND "FRK_EventDeliveryStore".Images[#Slot].Entries[#Position].Checksum = "FRK_DeliveryRowCrc"(Sequence := "FRK_EventDeliveryStore".Images[#Slot].Entries[#Position].Sequence, Ev := #Ev)
                AND (#Ev.State = 1 OR #Ev.State = 0)
                AND #Ev.ResetClass >= 0 AND #Ev.ResetClass <= 1
                AND #Ev.Severity >= 0 AND #Ev.Severity <= 2
                AND #Ev.Category >= 0 AND #Ev.Category <= 2
                AND #Ev.Description <> WSTRING#'' AND #Ev.SourcePath <> WSTRING#'' AND #Ev.Duration >= T#0ms;
            IF NOT #Valid THEN EXIT; END_IF;
            #Previous := "FRK_EventDeliveryStore".Images[#Slot].Entries[#Position].Sequence;
        END_FOR;
    END_IF;
    "FRK_EventDeliveryRuntime".Valid[#Slot] := #Valid;
    "FRK_DeliveryPublish"(Slot := #Slot);
END_FUNCTION

FUNCTION "FRK_DeliveryCapture" : Void
{ S7_Optimized_Access := 'TRUE' }
VERSION : 0.1
VAR_INPUT
    Ev : "ST_AlarmEvent";
END_VAR
VAR_IN_OUT
    AlarmLog : "FRK_AlarmLog";
END_VAR
VAR_TEMP
    Slot : Int;
    Position : Int;
END_VAR
BEGIN
    #Slot := #AlarmLog.DeliverySlot;
    IF #Slot < 1 OR #Slot > 1 OR #AlarmLog.DeliveryMuted THEN RETURN; END_IF;
    IF NOT "FRK_EventDeliveryRuntime".Valid[#Slot] THEN RETURN; END_IF;
    IF "FRK_EventDeliveryStore".Images[#Slot].Count >= 32 OR "FRK_EventDeliveryStore".Images[#Slot].NextSequence = UDINT#4294967295 THEN
        "FRK_EventDeliveryStore".Images[#Slot].Overflow := TRUE;
        IF "FRK_EventDeliveryStore".Images[#Slot].Dropped < UDINT#4294967295 THEN "FRK_EventDeliveryStore".Images[#Slot].Dropped := "FRK_EventDeliveryStore".Images[#Slot].Dropped + 1; END_IF;
        "FRK_DeliverySave"(Slot := #Slot);
        RETURN;
    END_IF;
    #Position := (("FRK_EventDeliveryStore".Images[#Slot].Head - 1 + "FRK_EventDeliveryStore".Images[#Slot].Count) MOD 32) + 1;
    "FRK_EventDeliveryStore".Images[#Slot].NextSequence := "FRK_EventDeliveryStore".Images[#Slot].NextSequence + 1;
    "FRK_EventDeliveryStore".Images[#Slot].Entries[#Position].Sequence := "FRK_EventDeliveryStore".Images[#Slot].NextSequence;
    "FRK_EventDeliveryStore".Images[#Slot].Entries[#Position].Ev := #Ev;
    "FRK_EventDeliveryStore".Images[#Slot].Entries[#Position].Checksum := "FRK_DeliveryRowCrc"(Sequence := "FRK_EventDeliveryStore".Images[#Slot].NextSequence, Ev := #Ev);
    "FRK_EventDeliveryStore".Images[#Slot].Count := "FRK_EventDeliveryStore".Images[#Slot].Count + 1;
    "FRK_DeliverySave"(Slot := #Slot);
END_FUNCTION

FUNCTION "FRK_DeliveryRequest" : Bool
{ S7_Optimized_Access := 'TRUE' }
VERSION : 0.1
VAR_INPUT
    RootScope : String;
    Request : "ST_HmiRequest";
    Access : "FRK_Access";
END_VAR
VAR_TEMP
    Slot : Int;
    Head : Int;
    Token : String[160];
    Prefix : String[254];
    Target : String[80];
END_VAR
BEGIN
    #FRK_DeliveryRequest := FALSE;
    // Receipts are data mutations, with a non-lowerable deployment minimum.
    IF #Access.CurrentLevel < 3 OR #Access.CurrentLevel < #Access.Policy.Required[1] THEN RETURN; END_IF;
    IF LEN(#Request.TargetPath) > 80 THEN RETURN; END_IF;
    #Target := WSTRING_TO_STRING(#Request.TargetPath);
    IF STRING_TO_WSTRING(#Target) <> #Request.TargetPath THEN RETURN; END_IF;
    #Prefix := CONCAT(IN1 := #RootScope, IN2 := '.');
    IF #Target <> #RootScope AND LEFT(IN := #Target, L := LEN(#Prefix)) <> #Prefix THEN RETURN; END_IF;
    #Slot := "FRK_DeliveryIndex"(Scope := #Target);
    IF #Slot < 1 OR #Slot > 1 THEN RETURN; END_IF;
    CASE #Request.Kind OF
        10001:
            IF NOT "FRK_EventDeliveryRuntime".Valid[#Slot] OR #Request.BoolValue THEN RETURN; END_IF;
            IF "FRK_EventDeliveryStore".Images[#Slot].Count <= 0 THEN RETURN; END_IF;
            #Head := "FRK_EventDeliveryStore".Images[#Slot].Head;
            IF #Head < 1 OR #Head > 32 THEN RETURN; END_IF;
            #Token := "FRK_DeliveryToken"(Slot := #Slot, Sequence := "FRK_EventDeliveryStore".Images[#Slot].Entries[#Head].Sequence);
            IF #Request.NameValue <> #Token OR #Request.DurationMs <> DWORD_TO_UDINT("FRK_EventDeliveryStore".Images[#Slot].Entries[#Head].Checksum) THEN RETURN; END_IF;
            "FRK_EventDeliveryStore".Images[#Slot].Entries[#Head].Sequence := 0;
            "FRK_EventDeliveryStore".Images[#Slot].Entries[#Head].Checksum := DWORD#0;
            "FRK_EventDeliveryStore".Images[#Slot].Entries[#Head].Ev := "FRK_UnitScratch".EmptyEvent;
            "FRK_EventDeliveryStore".Images[#Slot].Head := (#Head MOD 32) + 1;
            "FRK_EventDeliveryStore".Images[#Slot].Count := "FRK_EventDeliveryStore".Images[#Slot].Count - 1;
            "FRK_DeliverySave"(Slot := #Slot);
            #FRK_DeliveryRequest := TRUE;
        10002:
            IF "FRK_EventDeliveryRuntime".Valid[#Slot] OR NOT "FRK_EventDeliveryRuntime".AnchorValid[#Slot] OR NOT #Request.BoolValue THEN RETURN; END_IF;
            IF #Request.TextValue <> WSTRING#'6c62c9b6-57d9-41b5-b689-e0540f642b31' OR #Request.NameValue <> "FRK_DeliveryNumber"(Value := "FRK_EventDeliveryStore".Anchors[#Slot].Epoch)
                OR "FRK_EventDeliveryStore".Anchors[#Slot].Epoch = UDINT#4294967295 THEN RETURN; END_IF;
            // Advance the independently checked identity before discarding data.
            "FRK_EventDeliveryStore".Anchors[#Slot].Epoch := "FRK_EventDeliveryStore".Anchors[#Slot].Epoch + 1;
            "FRK_EventDeliveryStore".Anchors[#Slot].Checksum := "FRK_DeliveryAnchorCrc"(Slot := #Slot);
            "FRK_DeliveryInitialize"(Slot := #Slot, Discarded := TRUE);
            #FRK_DeliveryRequest := TRUE;
        ELSE RETURN;
    END_CASE;
END_FUNCTION

// Core section 7.7 prototype: private retained provider injection and independent root sessions.
// User records are salted Core-compatible hashes, never commissioning plaintext.
FUNCTION "FRK_Sha256Pin" : Bool
{ S7_Optimized_Access := 'TRUE' }
VERSION : 0.1
VAR_INPUT
    Size : DInt;
END_VAR
VAR_IN_OUT
    Data : Array[0..47] of Byte;
    Digest : Array[0..31] of Byte;
END_VAR
VAR_TEMP
    BlockBytes : Array[0..63] of Byte;
    Words : Array[0..63] of DWord;
    Hash : Array[0..7] of DWord;
    Index : DInt;
    A : DWord;
    B : DWord;
    C : DWord;
    D : DWord;
    E : DWord;
    F : DWord;
    G : DWord;
    H : DWord;
    S0 : DWord;
    S1 : DWord;
    T1 : DWord;
    T2 : DWord;
    K : Array[0..63] of DWord;
END_VAR
BEGIN
    #FRK_Sha256Pin := FALSE;
    #K[0] := DWORD#16#428A2F98;
    #K[1] := DWORD#16#71374491;
    #K[2] := DWORD#16#B5C0FBCF;
    #K[3] := DWORD#16#E9B5DBA5;
    #K[4] := DWORD#16#3956C25B;
    #K[5] := DWORD#16#59F111F1;
    #K[6] := DWORD#16#923F82A4;
    #K[7] := DWORD#16#AB1C5ED5;
    #K[8] := DWORD#16#D807AA98;
    #K[9] := DWORD#16#12835B01;
    #K[10] := DWORD#16#243185BE;
    #K[11] := DWORD#16#550C7DC3;
    #K[12] := DWORD#16#72BE5D74;
    #K[13] := DWORD#16#80DEB1FE;
    #K[14] := DWORD#16#9BDC06A7;
    #K[15] := DWORD#16#C19BF174;
    #K[16] := DWORD#16#E49B69C1;
    #K[17] := DWORD#16#EFBE4786;
    #K[18] := DWORD#16#0FC19DC6;
    #K[19] := DWORD#16#240CA1CC;
    #K[20] := DWORD#16#2DE92C6F;
    #K[21] := DWORD#16#4A7484AA;
    #K[22] := DWORD#16#5CB0A9DC;
    #K[23] := DWORD#16#76F988DA;
    #K[24] := DWORD#16#983E5152;
    #K[25] := DWORD#16#A831C66D;
    #K[26] := DWORD#16#B00327C8;
    #K[27] := DWORD#16#BF597FC7;
    #K[28] := DWORD#16#C6E00BF3;
    #K[29] := DWORD#16#D5A79147;
    #K[30] := DWORD#16#06CA6351;
    #K[31] := DWORD#16#14292967;
    #K[32] := DWORD#16#27B70A85;
    #K[33] := DWORD#16#2E1B2138;
    #K[34] := DWORD#16#4D2C6DFC;
    #K[35] := DWORD#16#53380D13;
    #K[36] := DWORD#16#650A7354;
    #K[37] := DWORD#16#766A0ABB;
    #K[38] := DWORD#16#81C2C92E;
    #K[39] := DWORD#16#92722C85;
    #K[40] := DWORD#16#A2BFE8A1;
    #K[41] := DWORD#16#A81A664B;
    #K[42] := DWORD#16#C24B8B70;
    #K[43] := DWORD#16#C76C51A3;
    #K[44] := DWORD#16#D192E819;
    #K[45] := DWORD#16#D6990624;
    #K[46] := DWORD#16#F40E3585;
    #K[47] := DWORD#16#106AA070;
    #K[48] := DWORD#16#19A4C116;
    #K[49] := DWORD#16#1E376C08;
    #K[50] := DWORD#16#2748774C;
    #K[51] := DWORD#16#34B0BCB5;
    #K[52] := DWORD#16#391C0CB3;
    #K[53] := DWORD#16#4ED8AA4A;
    #K[54] := DWORD#16#5B9CCA4F;
    #K[55] := DWORD#16#682E6FF3;
    #K[56] := DWORD#16#748F82EE;
    #K[57] := DWORD#16#78A5636F;
    #K[58] := DWORD#16#84C87814;
    #K[59] := DWORD#16#8CC70208;
    #K[60] := DWORD#16#90BEFFFA;
    #K[61] := DWORD#16#A4506CEB;
    #K[62] := DWORD#16#BEF9A3F7;
    #K[63] := DWORD#16#C67178F2;
    FOR #Index := 0 TO 31 DO #Digest[#Index] := 0; END_FOR;
    IF #Size < 0 OR #Size > 48 THEN RETURN; END_IF;
    // Authentication messages fit exactly one SHA-256 block.
    FOR #Index := 0 TO 63 DO #BlockBytes[#Index] := 0; END_FOR;
    FOR #Index := 0 TO #Size - 1 DO #BlockBytes[#Index] := #Data[#Index]; END_FOR;
    #BlockBytes[#Size] := BYTE#16#80;
    #BlockBytes[62] := DWORD_TO_BYTE(SHR(IN := DINT_TO_DWORD(#Size * 8), N := 8));
    #BlockBytes[63] := DINT_TO_BYTE(#Size * 8);
    #Hash[0] := DWORD#16#6A09E667;
    #Hash[1] := DWORD#16#BB67AE85;
    #Hash[2] := DWORD#16#3C6EF372;
    #Hash[3] := DWORD#16#A54FF53A;
    #Hash[4] := DWORD#16#510E527F;
    #Hash[5] := DWORD#16#9B05688C;
    #Hash[6] := DWORD#16#1F83D9AB;
    #Hash[7] := DWORD#16#5BE0CD19;
    FOR #Index := 0 TO 15 DO
        #Words[#Index] := SHL(IN := BYTE_TO_DWORD(#BlockBytes[4 * #Index]), N := 24)
            OR SHL(IN := BYTE_TO_DWORD(#BlockBytes[4 * #Index + 1]), N := 16)
            OR SHL(IN := BYTE_TO_DWORD(#BlockBytes[4 * #Index + 2]), N := 8)
            OR BYTE_TO_DWORD(#BlockBytes[4 * #Index + 3]);
    END_FOR;
    FOR #Index := 16 TO 63 DO
        #S0 := ROR(IN := #Words[#Index-15], N := 7) XOR ROR(IN := #Words[#Index-15], N := 18) XOR SHR(IN := #Words[#Index-15], N := 3);
        #S1 := ROR(IN := #Words[#Index-2], N := 17) XOR ROR(IN := #Words[#Index-2], N := 19) XOR SHR(IN := #Words[#Index-2], N := 10);
        #Words[#Index] := UDINT_TO_DWORD(ULINT_TO_UDINT(UDINT_TO_ULINT(DWORD_TO_UDINT(#Words[#Index-16])) + UDINT_TO_ULINT(DWORD_TO_UDINT(#S0)) + UDINT_TO_ULINT(DWORD_TO_UDINT(#Words[#Index-7])) + UDINT_TO_ULINT(DWORD_TO_UDINT(#S1))));
    END_FOR;
    #A := #Hash[0]; #B := #Hash[1]; #C := #Hash[2]; #D := #Hash[3];
    #E := #Hash[4]; #F := #Hash[5]; #G := #Hash[6]; #H := #Hash[7];
    FOR #Index := 0 TO 63 DO
        #S1 := ROR(IN := #E, N := 6) XOR ROR(IN := #E, N := 11) XOR ROR(IN := #E, N := 25);
        #T1 := UDINT_TO_DWORD(ULINT_TO_UDINT(UDINT_TO_ULINT(DWORD_TO_UDINT(#H)) + UDINT_TO_ULINT(DWORD_TO_UDINT(#S1)) + UDINT_TO_ULINT(DWORD_TO_UDINT((#E AND #F) XOR ((NOT #E) AND #G))) + UDINT_TO_ULINT(DWORD_TO_UDINT(#K[#Index])) + UDINT_TO_ULINT(DWORD_TO_UDINT(#Words[#Index]))));
        #S0 := ROR(IN := #A, N := 2) XOR ROR(IN := #A, N := 13) XOR ROR(IN := #A, N := 22);
        #T2 := UDINT_TO_DWORD(ULINT_TO_UDINT(UDINT_TO_ULINT(DWORD_TO_UDINT(#S0)) + UDINT_TO_ULINT(DWORD_TO_UDINT((#A AND #B) XOR (#A AND #C) XOR (#B AND #C)))));
        #H := #G; #G := #F; #F := #E;
        #E := UDINT_TO_DWORD(ULINT_TO_UDINT(UDINT_TO_ULINT(DWORD_TO_UDINT(#D)) + UDINT_TO_ULINT(DWORD_TO_UDINT(#T1))));
        #D := #C; #C := #B; #B := #A;
        #A := UDINT_TO_DWORD(ULINT_TO_UDINT(UDINT_TO_ULINT(DWORD_TO_UDINT(#T1)) + UDINT_TO_ULINT(DWORD_TO_UDINT(#T2))));
    END_FOR;
    #Words[0] := #A; #Words[1] := #B; #Words[2] := #C; #Words[3] := #D;
    #Words[4] := #E; #Words[5] := #F; #Words[6] := #G; #Words[7] := #H;
    FOR #Index := 0 TO 7 DO
        #Hash[#Index] := UDINT_TO_DWORD(ULINT_TO_UDINT(UDINT_TO_ULINT(DWORD_TO_UDINT(#Hash[#Index])) + UDINT_TO_ULINT(DWORD_TO_UDINT(#Words[#Index]))));
        #Digest[4 * #Index] := DWORD_TO_BYTE(SHR(IN := #Hash[#Index], N := 24));
        #Digest[4 * #Index + 1] := DWORD_TO_BYTE(SHR(IN := #Hash[#Index], N := 16));
        #Digest[4 * #Index + 2] := DWORD_TO_BYTE(SHR(IN := #Hash[#Index], N := 8));
        #Digest[4 * #Index + 3] := DWORD_TO_BYTE(#Hash[#Index]);
    END_FOR;
    FOR #Index := 0 TO 63 DO #BlockBytes[#Index] := 0; #Words[#Index] := 0; END_FOR;
    #FRK_Sha256Pin := TRUE;
END_FUNCTION

FUNCTION "FRK_AccessCancel" : Void
{ S7_Optimized_Access := 'TRUE' }
VERSION : 0.1
VAR_IN_OUT
    Access : "FRK_Access";
END_VAR
VAR_TEMP
    Index : DInt;
END_VAR
BEGIN
    #Access.LoginBusy := FALSE;
    #Access.CandidateUser := '';
    #Access.CandidateLevel := 0;
    #Access.Round := 0;
    FOR #Index := 0 TO 15 DO #Access.Salt[#Index] := 0; END_FOR;
    FOR #Index := 0 TO 31 DO #Access.Digest[#Index] := 0; #Access.Expected[#Index] := 0; END_FOR;
END_FUNCTION

FUNCTION "FRK_AccessLogout" : Void
{ S7_Optimized_Access := 'TRUE' }
VERSION : 0.1
VAR_IN_OUT
    Access : "FRK_Access";
END_VAR
BEGIN
    "FRK_AccessCancel"(Access := #Access);
    "FRK_AccessDropSession"(Access := #Access);
END_FUNCTION

FUNCTION "FRK_AccessDropSession" : Void
{ S7_Optimized_Access := 'TRUE' }
VERSION : 0.1
VAR_IN_OUT
    Access : "FRK_Access";
END_VAR
BEGIN
    #Access.CurrentLevel := 0;
    #Access.CurrentUser := '';
    #Access.LoginFailed := FALSE;
    #Access.SessionGeneration := "FRK_AccessNext"(Previous := #Access.SessionGeneration);
END_FUNCTION

FUNCTION "FRK_AccessNext" : UDInt
{ S7_Optimized_Access := 'TRUE' }
VERSION : 0.1
VAR_INPUT
    Previous : UDInt;
END_VAR
BEGIN
    IF #Previous = UDINT#4294967295 THEN #FRK_AccessNext := 1; ELSE #FRK_AccessNext := #Previous + 1; END_IF;
END_FUNCTION

FUNCTION "FRK_AccessLogin" : Void
{ S7_Optimized_Access := 'TRUE' }
VERSION : 0.1
VAR_INPUT
    User : String;
    Secret : String;
    Sequence : UDInt;
END_VAR
VAR_IN_OUT
    Access : "FRK_Access";
END_VAR
VAR_TEMP
    Data : Array[0..47] of Byte;
    Index : DInt;
    Slot : DInt;
    Size : Int;
    HashOk : Bool;
END_VAR
BEGIN
    "FRK_AccessCancel"(Access := #Access);
    #Access.LoginFailed := FALSE;
    #Access.LoginSequence := #Sequence;
    #Access.CandidateGeneration := "FRK_LocalUsers".Generation;
    #Access.LoginSince := "FRK_Clock".NowMs;
    #Access.LoginTimeoutMs := 6000;
    #Access.CandidateUser := #User;
    // Unknown users execute the same bounded work with a dummy salt/digest.
    IF #Access.ProviderEnabled AND "FRK_AccessStorage".UsersReady AND "FRK_LocalUsers".Count >= 0 AND "FRK_LocalUsers".Count <= 16 THEN
        FOR #Slot := 1 TO "FRK_LocalUsers".Count DO
            IF #User <> '' AND "FRK_LocalUsers".Rows[#Slot].User = #User THEN
                IF "FRK_LocalUsers".Rows[#Slot].Level >= 1 AND "FRK_LocalUsers".Rows[#Slot].Level <= 4 THEN
                    #Access.CandidateLevel := "FRK_LocalUsers".Rows[#Slot].Level;
                    #Access.Salt := "FRK_LocalUsers".Rows[#Slot].Salt;
                    #Access.Expected := "FRK_LocalUsers".Rows[#Slot].PinHash;
                END_IF;
                EXIT;
            END_IF;
        END_FOR;
    END_IF;
    FOR #Index := 0 TO 47 DO #Data[#Index] := 0; END_FOR;
    FOR #Index := 0 TO 15 DO #Data[#Index] := #Access.Salt[#Index]; END_FOR;
    #Size := LEN(#Secret);
    IF #Size > 32 THEN #Size := 0; #Access.CandidateLevel := 0; END_IF;
    FOR #Index := 1 TO #Size DO #Data[15 + #Index] := CHAR_TO_BYTE(#Secret[#Index]); END_FOR;
    #HashOk := "FRK_Sha256Pin"(Data := #Data, Size := 16 + INT_TO_DINT(#Size), Digest := #Access.Digest);
    FOR #Index := 0 TO 47 DO #Data[#Index] := 0; END_FOR;
    #Access.LoginBusy := #HashOk;
END_FUNCTION

FUNCTION "FRK_AccessAudit" : Void
{ S7_Optimized_Access := 'TRUE' }
VERSION : 0.1
VAR_INPUT
    What : WString;
    Who : String;
    SourcePath : WString;
END_VAR
VAR_IN_OUT
    AlarmLog : "FRK_AlarmLog";
END_VAR
VAR_TEMP
    Description : WString[480];
END_VAR
BEGIN
    #Description := CONCAT(IN1 := #What, IN2 := WSTRING#': ');
    #Description := CONCAT(IN1 := #Description, IN2 := STRING_TO_WSTRING(#Who));
    "FRK_AlarmMessage"(AlarmLog := #AlarmLog, Reason := 0, Description := #Description, SourcePath := #SourcePath);
END_FUNCTION

FUNCTION "FRK_AccessCyclic" : Void
{ S7_Optimized_Access := 'TRUE' }
VERSION : 0.1
VAR_INPUT
    Startup : Bool;
    SourcePath : WString;
END_VAR
VAR_IN_OUT
    Access : "FRK_Access";
    AlarmLog : "FRK_AlarmLog";
    Revision : UDInt;
END_VAR
VAR_TEMP
    Data : Array[0..47] of Byte;
    Index : DInt;
    Difference : Byte;
    HashOk : Bool;
END_VAR
BEGIN
    #Access.LoginTimeoutMs := 6000;
    IF #Startup THEN
        "FRK_AccessLogout"(Access := #Access);
        #Access.LoginResultSequence := 0;
    END_IF;
    IF #Access.ProviderGeneration <> "FRK_LocalUsers".Generation OR NOT "FRK_AccessStorage".UsersReady THEN
        IF #Access.CurrentLevel > 0 THEN
            "FRK_AccessAudit"(AlarmLog := #AlarmLog, What := WSTRING#'std.audit.autoLogout', Who := #Access.CurrentUser, SourcePath := #SourcePath);
            "FRK_AccessDropSession"(Access := #Access);
            #Revision := "FRK_ConfigRevision"(Previous := #Revision);
        END_IF;
        IF #Access.LoginBusy THEN #Access.CandidateLevel := 0; END_IF;
        #Access.ProviderGeneration := "FRK_LocalUsers".Generation;
    END_IF;
    IF #Access.CurrentLevel > 0 AND #Access.Policy.SessionTimeout > T#0ms THEN
        IF "FRK_Elapsed"(NewMs := "FRK_Clock".NowMs, OldMs := #Access.LastActivity) >= DINT_TO_UDINT(TIME_TO_DINT(#Access.Policy.SessionTimeout)) THEN
            "FRK_AccessAudit"(AlarmLog := #AlarmLog, What := WSTRING#'std.audit.autoLogout', Who := #Access.CurrentUser, SourcePath := #SourcePath);
            // Expiring the old session does not discard a separately committed
            // credential attempt. Explicit logout cancels both.
            "FRK_AccessDropSession"(Access := #Access);
            #Revision := "FRK_ConfigRevision"(Previous := #Revision);
        END_IF;
    END_IF;
    IF NOT #Access.LoginBusy THEN RETURN; END_IF;
    // One compression per active scan; never run all PIN rounds in one scan.
    FOR #Index := 0 TO 31 DO #Data[#Index] := #Access.Digest[#Index]; END_FOR;
    FOR #Index := 0 TO 15 DO #Data[32 + #Index] := #Access.Salt[#Index]; END_FOR;
    #HashOk := "FRK_Sha256Pin"(Data := #Data, Size := 48, Digest := #Access.Digest);
    FOR #Index := 0 TO 47 DO #Data[#Index] := 0; END_FOR;
    #Access.Round := #Access.Round + 1;
    IF NOT #HashOk OR "FRK_Elapsed"(NewMs := "FRK_Clock".NowMs, OldMs := #Access.LoginSince) >= #Access.LoginTimeoutMs THEN
        #Access.CandidateLevel := 0;
    ELSIF #Access.Round < 256 THEN RETURN;
    END_IF;
    #Difference := 0;
    FOR #Index := 0 TO 31 DO #Difference := #Difference OR (#Access.Digest[#Index] XOR #Access.Expected[#Index]); END_FOR;
    #Access.LoginFailed := #Difference <> 0 OR #Access.CandidateLevel = 0 OR NOT #Access.ProviderEnabled OR NOT "FRK_AccessStorage".UsersReady OR #Access.CandidateGeneration <> "FRK_LocalUsers".Generation;
    IF #Access.LoginFailed THEN
        "FRK_AccessAudit"(AlarmLog := #AlarmLog, What := WSTRING#'std.audit.loginFailed', Who := #Access.CandidateUser, SourcePath := #SourcePath);
    ELSE
        #Access.CurrentUser := #Access.CandidateUser;
        #Access.CurrentLevel := #Access.CandidateLevel;
        #Access.LastActivity := "FRK_Clock".NowMs;
        #Access.SessionGeneration := "FRK_AccessNext"(Previous := #Access.SessionGeneration);
        #Revision := "FRK_ConfigRevision"(Previous := #Revision);
        "FRK_AccessAudit"(AlarmLog := #AlarmLog, What := WSTRING#'std.audit.login', Who := #Access.CurrentUser, SourcePath := #SourcePath);
    END_IF;
    #Access.LoginResultSequence := #Access.LoginSequence;
    "FRK_AccessCancel"(Access := #Access);
END_FUNCTION

FUNCTION "FRK_AccessFinish" : Void
{ S7_Optimized_Access := 'TRUE' }
VERSION : 0.1
VAR_INPUT
    Unit : "FRK_Unit";
    Response : "ST_HmiResponse";
    SourcePath : WString;
END_VAR
VAR_IN_OUT
    Access : "FRK_Access";
    AlarmLog : "FRK_AlarmLog";
    Revision : UDInt;
END_VAR
VAR_TEMP
    What : WString[160];
    AuditPath : WString[255];
END_VAR
BEGIN
    IF NOT #Unit.RequestPending THEN RETURN; END_IF;
    CASE #Unit.Request.Kind OF
        23, 15,
        16, 17,
        1: RETURN;
        2:
            "FRK_AccessAudit"(AlarmLog := #AlarmLog, What := WSTRING#'std.audit.logout', Who := #Unit.RequestUser, SourcePath := #SourcePath);
            #Revision := "FRK_ConfigRevision"(Previous := #Revision);
            RETURN;
        ELSE #What := WSTRING#'std.audit.accessDenied';
    END_CASE;
    IF #Response.Accepted THEN
        #What := WSTRING#'std.audit.operatorAction';
        IF #Access.CurrentLevel > 0 THEN #Access.LastActivity := "FRK_Clock".NowMs; END_IF;
        IF #Unit.Request.Kind = 24 OR #Unit.Request.Kind = 25 THEN #Revision := "FRK_ConfigRevision"(Previous := #Revision); END_IF;
    END_IF;
    #AuditPath := #SourcePath;
    IF #Unit.Request.Kind = 11 THEN
        IF #Response.Accepted THEN #AuditPath := #Unit.Request.TargetPath; END_IF;
        IF #Response.Accepted THEN #What := WSTRING#'std.audit.manualCommandAccepted'; ELSE #What := WSTRING#'std.audit.manualCommandRejected'; END_IF;
    END_IF;
    #What := CONCAT(IN1 := #What, IN2 := WSTRING#' kind=');
    #What := CONCAT(IN1 := #What, IN2 := DINT_TO_WSTRING(#Unit.Request.Kind));
    #What := CONCAT(IN1 := #What, IN2 := WSTRING#' value=');
    #What := CONCAT(IN1 := #What, IN2 := DINT_TO_WSTRING(#Unit.Request.IntValue));
    "FRK_AccessAudit"(AlarmLog := #AlarmLog, What := #What, Who := #Unit.RequestUser, SourcePath := #AuditPath);
END_FUNCTION

// Canonical retained-image CRC primitives, shared by typed consumers.
FUNCTION "FRK_CrcByte" : DWord
{ S7_Optimized_Access := 'TRUE' }
VERSION : 0.1
VAR_INPUT
    Previous : DWord;
    Value : Byte;
END_VAR
VAR_TEMP
    BitIndex : Int;
    Work : DWord;
END_VAR
BEGIN
    #Work := #Previous XOR BYTE_TO_DWORD(#Value);
    FOR #BitIndex := 0 TO 7 DO
        IF (#Work AND DWORD#1) <> 0 THEN #Work := SHR(IN := #Work, N := 1) XOR DWORD#16#EDB88320;
        ELSE #Work := SHR(IN := #Work, N := 1); END_IF;
    END_FOR;
    #FRK_CrcByte := #Work;
END_FUNCTION

FUNCTION "FRK_CrcNumber" : DWord
{ S7_Optimized_Access := 'TRUE' }
VERSION : 0.1
VAR_INPUT
    Previous : DWord;
    Value : UDInt;
END_VAR
VAR_TEMP
    Index : Int;
    Work : DWord;
END_VAR
BEGIN
    #Work := #Previous;
    FOR #Index := 0 TO 3 DO
        #Work := "FRK_CrcByte"(Previous := #Work, Value := DWORD_TO_BYTE(SHR(IN := UDINT_TO_DWORD(#Value), N := INT_TO_UINT(#Index * 8))));
    END_FOR;
    #FRK_CrcNumber := #Work;
END_FUNCTION


// Reference-1500 LOCAL_RETAIN adapter. No sessions or plaintext credentials.
// CRC-32 arithmetic comes from Core F_Crc32; encoding is binding-local, versioned.
FUNCTION "FRK_AccessUsersCrc" : DWord
{ S7_Optimized_Access := 'TRUE' }
VERSION : 0.1
VAR_TEMP
    Work : DWord;
    Slot : Int;
    Index : Int;
    Size : Int;
END_VAR
BEGIN
    #Work := "FRK_CrcNumber"(Previous := DWORD#16#FFFFFFFF, Value := UINT_TO_UDINT("FRK_LocalUsers".SchemaVersion));
    #Work := "FRK_CrcNumber"(Previous := #Work, Value := "FRK_LocalUsers".Generation);
    #Work := "FRK_CrcNumber"(Previous := #Work, Value := DINT_TO_UDINT("FRK_LocalUsers".Count));
    // Unused rows are included: an altered dormant credential is not ignored.
    FOR #Slot := 1 TO 16 DO
        #Size := LEN("FRK_LocalUsers".Rows[#Slot].User);
        #Work := "FRK_CrcNumber"(Previous := #Work, Value := INT_TO_UDINT(#Size));
        FOR #Index := 1 TO #Size DO
            #Work := "FRK_CrcByte"(Previous := #Work, Value := CHAR_TO_BYTE("FRK_LocalUsers".Rows[#Slot].User[#Index]));
        END_FOR;
        #Work := "FRK_CrcNumber"(Previous := #Work, Value := DINT_TO_UDINT("FRK_LocalUsers".Rows[#Slot].Level));
        FOR #Index := 0 TO 15 DO
            #Work := "FRK_CrcByte"(Previous := #Work, Value := "FRK_LocalUsers".Rows[#Slot].Salt[#Index]);
        END_FOR;
        FOR #Index := 0 TO 31 DO
            #Work := "FRK_CrcByte"(Previous := #Work, Value := "FRK_LocalUsers".Rows[#Slot].PinHash[#Index]);
        END_FOR;
    END_FOR;
    #FRK_AccessUsersCrc := NOT #Work;
END_FUNCTION

FUNCTION "FRK_AccessUsersShape" : Bool
{ S7_Optimized_Access := 'TRUE' }
VERSION : 0.1
VAR_TEMP
    Slot : Int;
    Other : Int;
END_VAR
BEGIN
    #FRK_AccessUsersShape := FALSE;
    IF "FRK_LocalUsers".Count < 0 OR "FRK_LocalUsers".Count > 16 THEN RETURN; END_IF;
    FOR #Slot := 1 TO DINT_TO_INT("FRK_LocalUsers".Count) DO
        IF "FRK_LocalUsers".Rows[#Slot].User = '' OR "FRK_LocalUsers".Rows[#Slot].Level < 0 OR "FRK_LocalUsers".Rows[#Slot].Level > 4 THEN RETURN; END_IF;
        FOR #Other := 1 TO #Slot - 1 DO
            IF "FRK_LocalUsers".Rows[#Slot].User = "FRK_LocalUsers".Rows[#Other].User THEN RETURN; END_IF;
        END_FOR;
    END_FOR;
    #FRK_AccessUsersShape := TRUE;
END_FUNCTION

FUNCTION "FRK_AccessUsersCommit" : Bool
{ S7_Optimized_Access := 'TRUE' }
VERSION : 0.1
BEGIN
    #FRK_AccessUsersCommit := "FRK_AccessUsersShape"();
    IF NOT #FRK_AccessUsersCommit THEN RETURN; END_IF;
    "FRK_LocalUsers".SchemaVersion := 1;
    "FRK_LocalUsers".Generation := "FRK_AccessNext"(Previous := "FRK_LocalUsers".Generation);
    "FRK_LocalUsers".Checksum := "FRK_AccessUsersCrc"();
    "FRK_AccessStorage".UsersCommissioned := TRUE;
    "FRK_AccessStorage".UsersReady := TRUE;
    "FRK_AccessStorage".UsersLost := FALSE;
END_FUNCTION

FUNCTION "FRK_AccessRegisterHash" : Bool
{ S7_Optimized_Access := 'TRUE' }
VERSION : 0.1
VAR_INPUT
    Record : "ST_UserRecord";
END_VAR
VAR_TEMP
    Slot : Int;
    Index : Int;
END_VAR
BEGIN
    // Trusted composition/provider seam, never a remote credential editor.
    #FRK_AccessRegisterHash := FALSE;
    IF NOT "FRK_AccessStorage".UsersReady OR #Record.User = '' OR #Record.Level < 0 OR #Record.Level > 4 THEN RETURN; END_IF;
    #Slot := 0;
    FOR #Index := 1 TO DINT_TO_INT("FRK_LocalUsers".Count) DO
        IF "FRK_LocalUsers".Rows[#Index].User = #Record.User THEN #Slot := #Index; EXIT; END_IF;
    END_FOR;
    IF #Slot = 0 THEN
        IF "FRK_LocalUsers".Count = 16 THEN RETURN; END_IF;
        "FRK_LocalUsers".Count := "FRK_LocalUsers".Count + 1;
        #Slot := DINT_TO_INT("FRK_LocalUsers".Count);
    END_IF;
    "FRK_LocalUsers".Rows[#Slot] := #Record;
    #FRK_AccessRegisterHash := "FRK_AccessUsersCommit"();
END_FUNCTION

FUNCTION "FRK_AccessStoreBoot" : Void
{ S7_Optimized_Access := 'TRUE' }
VERSION : 0.1
VAR_INPUT
    Startup : Bool;
END_VAR
VAR_TEMP
    Accepted : Bool;
END_VAR
BEGIN
    IF NOT #Startup THEN RETURN; END_IF;
    "FRK_AccessStorage".UsersReady := FALSE;
    "FRK_AccessStorage".UsersLost := FALSE;
    // A virgin image may accept deliberate composition-root provisioning.
    IF NOT "FRK_AccessStorage".UsersCommissioned AND "FRK_LocalUsers".SchemaVersion = 0 AND "FRK_LocalUsers".Generation = 0 AND "FRK_LocalUsers".Checksum = DWORD#0 THEN
        #Accepted := "FRK_AccessUsersCommit"();
        "FRK_AccessStorage".UsersLost := NOT #Accepted;
    ELSIF "FRK_AccessStorage".UsersCommissioned AND "FRK_LocalUsers".SchemaVersion = 1 AND "FRK_LocalUsers".Generation > 0 AND "FRK_AccessUsersShape"() THEN
        "FRK_AccessStorage".UsersReady := "FRK_LocalUsers".Checksum = "FRK_AccessUsersCrc"();
        "FRK_AccessStorage".UsersLost := NOT "FRK_AccessStorage".UsersReady;
    ELSE "FRK_AccessStorage".UsersLost := TRUE;
    END_IF;
END_FUNCTION

FUNCTION "FRK_AccessPolicyCrc" : DWord
{ S7_Optimized_Access := 'TRUE' }
VERSION : 0.1
VAR_IN_OUT
    Image : "FRK_AccessPolicyImage";
END_VAR
VAR_TEMP
    Work : DWord;
    Index : Int;
    Size : Int;
END_VAR
BEGIN
    #Work := "FRK_CrcNumber"(Previous := DWORD#16#FFFFFFFF, Value := UINT_TO_UDINT(#Image.SchemaVersion));
    IF #Image.Initialized THEN #Work := "FRK_CrcByte"(Previous := #Work, Value := BYTE#1);
    ELSE #Work := "FRK_CrcByte"(Previous := #Work, Value := BYTE#0); END_IF;
    #Work := "FRK_CrcNumber"(Previous := #Work, Value := #Image.Generation);
    #Size := LEN(#Image.Scope);
    #Work := "FRK_CrcNumber"(Previous := #Work, Value := INT_TO_UDINT(#Size));
    FOR #Index := 1 TO #Size DO #Work := "FRK_CrcByte"(Previous := #Work, Value := CHAR_TO_BYTE(#Image.Scope[#Index])); END_FOR;
    FOR #Index := 0 TO 11 DO
        #Work := "FRK_CrcNumber"(Previous := #Work, Value := DINT_TO_UDINT(#Image.Policy.Required[#Index]));
    END_FOR;
    #Work := "FRK_CrcNumber"(Previous := #Work, Value := DINT_TO_UDINT(TIME_TO_DINT(#Image.Policy.SessionTimeout)));
    #FRK_AccessPolicyCrc := NOT #Work;
END_FUNCTION

FUNCTION "FRK_AccessPolicyShape" : Bool
{ S7_Optimized_Access := 'TRUE' }
VERSION : 0.1
VAR_IN_OUT
    Policy : "ST_AccessPolicy";
END_VAR
VAR_TEMP
    Index : Int;
END_VAR
BEGIN
    #FRK_AccessPolicyShape := FALSE;
    IF #Policy.SessionTimeout < T#0ms OR #Policy.SessionTimeout > T#604800000ms THEN RETURN; END_IF;
    FOR #Index := 0 TO 11 DO
        IF #Policy.Required[#Index] < 0 OR #Policy.Required[#Index] > 4 THEN RETURN; END_IF;
    END_FOR;
    #FRK_AccessPolicyShape := TRUE;
END_FUNCTION

FUNCTION "FRK_AccessPolicyValid" : Bool
{ S7_Optimized_Access := 'TRUE' }
VERSION : 0.1
VAR_IN_OUT
    Image : "FRK_AccessPolicyImage";
END_VAR
VAR_TEMP
    Index : Int;
END_VAR
BEGIN
    #FRK_AccessPolicyValid := FALSE;
    IF NOT #Image.Initialized OR #Image.SchemaVersion <> 1 OR #Image.Scope = '' OR #Image.Generation = 0 OR NOT "FRK_AccessPolicyShape"(Policy := #Image.Policy) THEN RETURN; END_IF;
    #FRK_AccessPolicyValid := #Image.Checksum = "FRK_AccessPolicyCrc"(Image := #Image);
END_FUNCTION

FUNCTION "FRK_AccessPolicySave" : Void
{ S7_Optimized_Access := 'TRUE' }
VERSION : 0.1
VAR_INPUT
    Scope : String;
END_VAR
VAR_IN_OUT
    Access : "FRK_Access";
END_VAR
BEGIN
    IF #Access.PolicySlot < 1 OR #Access.PolicySlot > 1 THEN RETURN; END_IF;
    IF #Scope = '' OR NOT "FRK_AccessPolicyShape"(Policy := #Access.Policy) THEN #Access.PolicyLost := TRUE; RETURN; END_IF;
    "FRK_AccessPolicies".Rows[#Access.PolicySlot].SchemaVersion := 1;
    "FRK_AccessPolicies".Rows[#Access.PolicySlot].Initialized := TRUE;
    "FRK_AccessPolicies".Rows[#Access.PolicySlot].Scope := #Scope;
    "FRK_AccessPolicies".Rows[#Access.PolicySlot].Generation := "FRK_AccessNext"(Previous := "FRK_AccessPolicies".Rows[#Access.PolicySlot].Generation);
    "FRK_AccessPolicies".Rows[#Access.PolicySlot].Policy := #Access.Policy;
    "FRK_AccessPolicies".Rows[#Access.PolicySlot].Checksum := "FRK_AccessPolicyCrc"(Image := "FRK_AccessPolicies".Rows[#Access.PolicySlot]);
END_FUNCTION

FUNCTION "FRK_AccessPolicyBoot" : Void
{ S7_Optimized_Access := 'TRUE' }
VERSION : 0.1
VAR_INPUT
    Startup : Bool;
    Root : Bool;
    Scope : String;
END_VAR
VAR_IN_OUT
    Access : "FRK_Access";
END_VAR
VAR_TEMP
    Index : Int;
    FreeSlot : Int;
END_VAR
BEGIN
    IF NOT #Startup THEN RETURN; END_IF;
    #Access.PolicySlot := 0; #Access.PolicyLost := FALSE;
    #Access.PolicyLossAlarm := 0; #Access.UserLossAlarm := 0;
    IF NOT #Root THEN RETURN; END_IF;
    #FreeSlot := 0;
    FOR #Index := 1 TO 1 DO
        IF "FRK_AccessPolicies".Rows[#Index].Scope = #Scope THEN
            IF #Access.PolicySlot <> 0 THEN #Access.PolicyLost := TRUE;
            ELSE #Access.PolicySlot := #Index; END_IF;
        ELSIF #FreeSlot = 0 AND NOT "FRK_AccessPolicies".Rows[#Index].Initialized AND "FRK_AccessPolicies".Rows[#Index].Scope = '' AND "FRK_AccessPolicies".Rows[#Index].SchemaVersion = 0 AND "FRK_AccessPolicies".Rows[#Index].Generation = 0 AND "FRK_AccessPolicies".Rows[#Index].Checksum = DWORD#0 THEN
            #FreeSlot := #Index;
        END_IF;
    END_FOR;
    IF #Access.PolicySlot > 0 THEN
        IF NOT #Access.PolicyLost AND "FRK_AccessPolicyValid"(Image := "FRK_AccessPolicies".Rows[#Access.PolicySlot]) THEN
            #Access.Policy := "FRK_AccessPolicies".Rows[#Access.PolicySlot].Policy;
        ELSE #Access.PolicyLost := TRUE;
        END_IF;
    ELSIF #FreeSlot > 0 THEN
        #Access.PolicySlot := #FreeSlot;
        "FRK_AccessPolicySave"(Access := #Access, Scope := #Scope);
    ELSE #Access.PolicyLost := TRUE;
    END_IF;
    IF #Access.PolicyLost THEN
        // Do not silently reopen actions after losing commissioned policy.
        #Access.Policy := "FRK_AccessStorage".EmptyPolicy;
        FOR #Index := 0 TO 11 DO #Access.Policy.Required[#Index] := 4; END_FOR;
    END_IF;
END_FUNCTION

